(* IEC 61131-3 sources: daoli-st-library/DL_Algo (part 5) *)

(* ---- FC_DL_DewPointCalc.st ---- *)
(*==============================================================================
 * 组件名称 (Component)  : FC_DL_DewPointCalc
 * 所属子库 (Sublibrary) : DL_Algo
 * 当前版本 (Version)    : 1.0.1
 * 兼容性   (Platform)   : CODESYS 3.5 / TwinCAT 3 / 汇川 InoProShop / Machine Expert
 *                         仅依赖 Standard.library（LN / EXP / ABS / MIN / MAX），
 *                         零厂商方言
 * 功能描述 (Function)   : Magnus-Tetens（Stull 参数化）露点温度计算。由干球
 *                         温度与相对湿度求露点：gamma := LN(RH/100) +
 *                         a*T/(b+T)，Td := b*gamma/(a-gamma)，a=17.625、
 *                         b=243.04（过水面参数化）。另附实际水汽压输出供
 *                         焓值类组件复用。现场用途：洁净室 / 干燥房环控、
 *                         冷面结露风险判断（表面温度低于露点即结露）。
 * 开源溯源 (Origin)     : 原创实现。公式为公开气象学 Magnus-Tetens/Stull
 *                         参数化（clean-room），按本库故障码体系重写并加严。
 * 属主转移 (R23 裁定)   : Magnus-Tetens 常数（a=17.625、b=243.04）唯一属主
 *                         自 R23 起为 FC_DL_VaporPressureSat；本件内联常数
 *                         为属主口径的历史引用，本版仅声明、逻辑零改动，
 *                         后续口径变更以属主件为单一事实源。
 * 设计验证 (Verified)   : python 6 位小数核验（a=17.625、b=243.04）：
 *                         T=25.0 度 RH=60.0 -> Td=16.698 度（约 16.7 达标）；
 *                         T=0.0 度 RH=100.0 -> Td=0.000 度（精确归零）；
 *                         T=20.0 度 RH=50.0 -> Td=9.261 度；
 *                         T=25.0 度 RH=60.0 -> fVaporPa=1897.8 Pa。
 * 验收向量 (Acceptance) :
 *   V1 T=25.0 RH=60.0：返回值约 16.698（容差 0.3），fVaporPa 约 1897.8
 *   V2 T=0.0 RH=100.0：返回值 0.000（容差 1E-3），uErrorId=0
 *   V3 T=20.0 RH=50.0：返回值约 9.261（容差 0.3）
 *   V4 RH=0.0：钳位至 0.1，uErrorId=16#0002_1501，返回确定值不发散
 *   V5 T=100.0：钳位至 60.0，uErrorId=16#0002_1502，bInRange=FALSE
 *   V6 T=-500.0：钳位至 -40.0，返回哨兵口径确定值，绝不返回未初始化值
 *   V7 RH=0.0：钳位至 0.1，LN 输入恒正不发散，返回值有限且为确定数
 *   V8 T=25.0 RH=60.0：fVaporPa 约 1897.8 Pa（容差 5.0），供焓值链路复用
 * 依赖     (Depends)    : 无 DL_ 内部依赖；仅标准 LN / EXP
 * 红线自检 (Redline)    : R1 ✓ 零全局变量表与外部变量引用 ｜ R2 ✓ 零物理 IO 地址直写
 *                         R3 ✓ 纯 IEC 61131-3 ｜ R4 ✓ 钳位+容差+防除零+出口默认值
 *                         R5 ✓ 全变量中英双语同行注释 ｜ R6 N/A（FC 无状态机）
 *                         R7 N/A（无实例调用）
 * 无状态声明 (Stateless): FC 全程无隐式状态，同输入必得同输出；
 *                         除 VAR_IN_OUT 之外的隐式状态为零。
 * 修订历史 (Revision)   :
 *   2026-11-15  v1.0.0  首版入库（Round 04 · Phase 3 · DL_Algo 批次）
 *============================================================================*)

(*-----------------------------------------------------------------------------
 * 调用示例 (Instance guide)：
 *   fTd := FC_DL_DewPointCalc(fTempC := stAir.fTemp,
 *                             fRhPct := stAir.fRh,
 *                             uErrorId => uDewErr,
 *                             fVaporPa => fVp,
 *                             bInRange => bInDom);
 *   结露联锁判定：IF (stChiller.fSurfTemp <= fTd) THEN bCondenseRisk := TRUE;
 *   注意：仅当 uErrorId = 0 且 bInRange = TRUE 时才可将 fTd 用于联锁判断。
 *   多测点批量换算：每个温湿度测点独立调用一次，函数无状态可安全复用。
 *   哨兵口径复核：任何返回值等于 -40.0 时必须先核对 uErrorId 再使用。
 *----------------------------------------------------------------------------*)

(*-----------------------------------------------------------------------------
 * 常见误用与现场提示 (Field notes)：
 *   1 湿度给成绝对湿度或露点值会得到荒谬结果，本函数只接收相对湿度百分数。
 *   2 冰点以下本函数按过水面参数化计算霜点近似值，误差略增，精密工艺
 *     场景（如锂电干燥房露点仪对标）建议上层做冰面 Magnus 修正。
 *   3 返回哨兵值 -40.0 仅为异常路径确定值口径，不构成有效露点数据，
 *     上位趋势画面应按 uErrorId 过滤后再绘图。
 *   4 本函数每周期都可调用，纯计算无副作用可放心放入高速任务；
 *     但输入应来自滤波后的温湿度信号，露点输出抖动会带抖联锁逻辑。
 *   5 fVaporPa 与露点同源同口径，做焓值或含湿量换算时无需二次查表，
 *     避免两套公式口径漂移导致热平衡算不平。
 *----------------------------------------------------------------------------*)
FUNCTION FC_DL_DewPointCalc : REAL
VAR_INPUT
    fTempC  : REAL;                      // 干球温度 [摄氏度]，有效域 -40..60 / Dry-bulb temperature [degC], valid range -40..60
    fRhPct  : REAL;                      // 相对湿度 [百分数]，有效域 0.1..100 / Relative humidity [percent], valid range 0.1..100
END_VAR
VAR_OUTPUT
    uErrorId : UDINT;                    // 故障码，0 = 无故障 / Error code, 0 = no error
    fVaporPa : REAL;                     // 实际水汽压 [Pa]，诊断与焓值复用 / Actual vapor pressure [Pa], diagnostic and reuse
    bInRange : BOOL;                     // 输入是否处于公式有效域 / Whether inputs are within the formula valid domain
END_VAR
VAR
    fGamma   : REAL;                     // Magnus 中间量 [1] / Magnus intermediate value [1]
    fRhEff   : REAL;                     // 钳位后的生效湿度 [百分数] / Effective clamped humidity [percent]
    fTempEff : REAL;                     // 钳位后的生效温度 [摄氏度] / Effective clamped temperature [degC]
END_VAR
VAR CONSTANT
    DL_DEW_A      : REAL := 17.625;      // Magnus 系数 a [1] / Magnus coefficient a [1]
    DL_DEW_C      : REAL := 243.04;      // Magnus 系数 b [摄氏度] / Magnus coefficient b [degC]
    DL_DEW_E0     : REAL := 611.2;       // 0 摄氏度饱和水汽压 [Pa] / Saturation vapor pressure at 0 degC [Pa]
    DL_DEW_T_MIN  : REAL := -40.0;       // 温度有效域下限 [摄氏度] / Temperature valid range low [degC]
    DL_DEW_T_MAX  : REAL := 60.0;        // 温度有效域上限 [摄氏度] / Temperature valid range high [degC]
    DL_DEW_RH_MIN : REAL := 0.1;         // 湿度工程下限 [百分数]，防对数发散 / Humidity engineering floor [percent], guards log divergence
    DL_DEW_SENTINEL : REAL := -40.0;     // 异常路径返回哨兵值 [摄氏度] / Sentinel return on error paths [degC]
    DL_DEW_EPS    : REAL := 1.0E-6;      // 浮点判零容差 / Float zero tolerance
    DL_DEW_INF_MAX : REAL := 1.0E30;     // 有限值判定幅值上限 / Magnitude bound for finite-value check
END_VAR

(*------------------------------------------------------------------------------
 * 段 1｜出口默认值（IEC 61131-3 强制）：入口即赋确定值，任何提前 RETURN
 *      前输出已确定；异常路径返回哨兵值 -40.0（安全下限口径）
 *      Exit defaults (mandatory): outputs assigned deterministically on entry
 *-----------------------------------------------------------------------------*)
FC_DL_DewPointCalc := DL_DEW_SENTINEL;               // 返回值哨兵预置 / Return value preset to sentinel
uErrorId           := 16#0002_0000;                  // 故障码先清零 / Error code cleared first
fVaporPa           := 0.0;                           // 水汽压默认置零 / Vapor pressure defaulted to zero
bInRange           := TRUE;                          // 默认视为在有效域 / Default considered in valid domain
fRhEff             := DL_DEW_RH_MIN;                 // 湿度预置工程下限 / Humidity preset to engineering floor
fTempEff           := DL_DEW_T_MIN;                  // 温度预置域下限 / Temperature preset to domain floor

(*------------------------------------------------------------------------------
 * 段 2｜非有限值防御：NaN 或超幅值输入直接返回哨兵并置公共码
 *      Non-finite defense: NaN or over-range input returns sentinel with code
 *-----------------------------------------------------------------------------*)
IF (fTempC <> fTempC) OR (ABS(fTempC) > DL_DEW_INF_MAX)
   OR (fRhPct <> fRhPct) OR (ABS(fRhPct) > DL_DEW_INF_MAX) THEN
    uErrorId           := 16#0002_0004;               // 输入非有限值已拒绝 / Non-finite input rejected
    FC_DL_DewPointCalc := DL_DEW_SENTINEL;
    fVaporPa           := 0.0;
    bInRange           := FALSE;
    RETURN;
END_IF

(*------------------------------------------------------------------------------
 * 段 3｜湿度钳位：下限防 LN(0) 发散，上限防超饱和非物理输入
 *      Humidity clamping: floor guards log divergence, cap blocks supersaturation
 *-----------------------------------------------------------------------------*)
IF fRhPct < DL_DEW_RH_MIN THEN
    fRhEff   := DL_DEW_RH_MIN;                       // 过低湿度钳位到工程下限 / Too low humidity clamped to floor
    uErrorId := 16#0002_1501;                        // 湿度越界已钳位 / Humidity out of range clamped
ELSIF fRhPct > 100.0 THEN
    fRhEff   := 100.0;                               // 超饱和湿度钳位到 100 / Supersaturated humidity clamped to 100
    uErrorId := 16#0002_1501;                        // 湿度越界已钳位 / Humidity out of range clamped
ELSE
    fRhEff := fRhPct;                                // 合法湿度原值生效 / Valid humidity applied as-is
END_IF

(*------------------------------------------------------------------------------
 * 段 4｜温度钳位：越域修正并标记不在有效域（含冰面霜点未计算提示口径）
 *      Temperature clamping: out-of-domain corrected and flagged
 *-----------------------------------------------------------------------------*)
IF (fTempC < DL_DEW_T_MIN) OR (fTempC > DL_DEW_T_MAX) THEN
    fTempEff := MIN(MAX(fTempC, DL_DEW_T_MIN), DL_DEW_T_MAX); // 双侧钳位到有效域 / Two-sided clamp into valid range
    uErrorId := 16#0002_1502;                        // 温度越域已钳位 / Temperature out of domain clamped
    bInRange := FALSE;                               // 标记不在公式有效域 / Flagged outside formula valid domain
ELSE
    fTempEff := fTempC;                              // 合法温度原值生效 / Valid temperature applied as-is
END_IF

(*------------------------------------------------------------------------------
 * 段 5｜分母防御性双检：b+fTempEff 理论上恒大于零（T>=-40），仍强制校验
 *      Defensive double check on denominator, theoretically always positive
 *-----------------------------------------------------------------------------*)
IF ABS(DL_DEW_C + fTempEff) <= DL_DEW_EPS THEN
    uErrorId           := 16#0002_1502;               // 分母异常按温度类故障处理 / Denominator anomaly treated as temperature fault
    FC_DL_DewPointCalc := DL_DEW_SENTINEL;
    fVaporPa           := 0.0;
    bInRange           := FALSE;
    RETURN;
END_IF

(*------------------------------------------------------------------------------
 * 段 6｜Magnus-Tetens 主体计算：gamma 中间量 + 露点反解 + 水汽压
 *      Magnus-Tetens core: gamma intermediate, dew point inversion, vapor pressure
 *      LN 输入恒大于零由湿度工程下限 0.1 保证，无需再判
 *      gamma 物理含义：对数形式的水汽分压与饱和分压比值度量，
 *      温度越高、湿度越大 gamma 越大，露点随之单调上移
 *-----------------------------------------------------------------------------*)
fGamma := LN(fRhEff / 100.0) + DL_DEW_A * fTempEff / (DL_DEW_C + fTempEff); // Magnus 中间量 / Magnus intermediate value

(* 分母 a-gamma：露点反解系数，由 gamma 单调有界性保证远离零，仍双检 *)
(* Denominator a-gamma: bounded away from zero by monotonicity, still guarded *)
IF ABS(DL_DEW_A - fGamma) <= DL_DEW_EPS THEN
    uErrorId           := 16#0002_1502;               // 反解分母异常按温度类故障处理 / Inversion denominator anomaly
    FC_DL_DewPointCalc := DL_DEW_SENTINEL;
    fVaporPa           := 0.0;
    bInRange           := FALSE;
    RETURN;
END_IF

FC_DL_DewPointCalc := DL_DEW_C * fGamma / (DL_DEW_A - fGamma); // 露点温度 [摄氏度] / Dew point temperature [degC]

(* 实际水汽压：饱和水汽压按当前温度指数外推后乘以相对湿度份额 *)
(* Actual vapor pressure: saturation pressure extrapolated by temperature times RH share *)
fVaporPa := DL_DEW_E0 * EXP(DL_DEW_A * fTempEff / (DL_DEW_C + fTempEff)) * fRhEff / 100.0;
END_FUNCTION

(* ---- FC_DL_DiverterLeadTimeCalc.st ---- *)
(*
  DL Factory R83 | FC_DL_DiverterLeadTimeCalc
  功能：按执行机构动作时间与线速算分流器提前量，反算触发延时并判可实现性。
  开源溯源：无（clean-room 自研，依据公开工艺公式，来源=行业通用公式，许可证=MIT，借鉴点=公式结构）
  规则：R1-R21 全遵守
*)
FUNCTION FC_DL_DiverterLeadTimeCalc : REAL
VAR_INPUT
    fConvSpeedMps   : REAL; // 输送线速度 [m/s] / Conveyor speed [m/s]
    fActuatorMs     : REAL; // 分流器全行程动作时间 [ms] / Diverter full-stroke time [ms]
    fSensorToPivotM : REAL; // 检测位到分流点距离 [m] / Sensor-to-pivot distance [m]
    fItemLenM       : REAL; // 物件长度 [m] / Item length along travel [m]
END_VAR
VAR_OUTPUT
    fLeadM          : REAL; // 需提前动作的等效距离 [m] / Required lead distance [m]
    fTriggerDelayMs : REAL; // 从检测沿到发出动作指令的延时 [ms] / Trigger delay after sensor edge [ms]
    xFeasible       : BOOL; // 时序可实现（延时非负且不超总输送时间）/ Timing feasible flag
    xValid          : BOOL; // 计算有效性标志 / Calculation validity flag
END_VAR
VAR
    fTotalMs : REAL; // 检测位到分流点总输送时间 [ms] / Total transit time [ms]
END_VAR
// 出口预置：四出口统一预置，可实现标志预置 FALSE（安全侧）
fLeadM := 0.0; fTriggerDelayMs := 0.0; xFeasible := FALSE; xValid := FALSE;
// 非有限拦截 + 量纲自检 + 速度零闸（R4/R20/R21）
IF NOT (fConvSpeedMps > -1.0E30 AND fConvSpeedMps < 1.0E30) OR NOT (fActuatorMs > -1.0E30 AND fActuatorMs < 1.0E30) OR NOT (fSensorToPivotM > -1.0E30 AND fSensorToPivotM < 1.0E30) OR NOT (fItemLenM > -1.0E30 AND fItemLenM < 1.0E30) OR fConvSpeedMps <= 0.0 OR fActuatorMs < 0.0 OR fSensorToPivotM <= 0.0 OR fItemLenM < 0.0 THEN
    FC_DL_DiverterLeadTimeCalc := -1.0; RETURN;   // 哨兵 -1：非有限或量纲越界 / Sentinel -1
END_IF
// 提前量：线速 × 动作时间(s) + 半件长（使物件中心对准分流点），m/s × s = m
fLeadM := fConvSpeedMps * (fActuatorMs / 1000.0) + fItemLenM / 2.0; // 提前量 [m] / Lead distance [m]
// 总输送时间：m ÷ (m/s) = s，×1000 = ms（分母已判正）
fTotalMs := (fSensorToPivotM / fConvSpeedMps) * 1000.0;   // 总输送时间 [ms] / Total transit time [ms]
// 触发延时：总输送时间 - 提前量对应时间（m ÷ m/s × 1000 = ms，量纲自洽）
fTriggerDelayMs := fTotalMs - (fLeadM / fConvSpeedMps) * 1000.0; // 触发延时 [ms] / Trigger delay [ms]
// 可实现性闸：负延时=前置距离不足；延时超总时间=参数逻辑倒置
IF fTriggerDelayMs < 0.0 THEN
    fTriggerDelayMs := 0.0;         // 负延时钳零（立即动作）/ Negative delay clamped, act at once
    xFeasible       := FALSE;       // 前置距离不足，不可分拣 / Insufficient lead distance
    xValid          := TRUE;        // 计算有效，仅结论不可行 / Calculation valid, conclusion infeasible
ELSIF fTriggerDelayMs <= fTotalMs THEN
    xFeasible := TRUE;              // 时序可实现 / Timing feasible
    xValid    := TRUE;              // 链路有效 / Chain valid
ELSE
    fTriggerDelayMs := fTotalMs;    // 延时超总时间钳位 / Clamp delay to total transit
    xFeasible       := FALSE;       // 逻辑倒置判不可行 / Inverted logic flagged
    xValid          := FALSE;       // 参数异常 / Parameter anomaly
END_IF
FC_DL_DiverterLeadTimeCalc := fTriggerDelayMs; // 返回触发延时 [ms] / Return trigger delay [ms]
END_FUNCTION

(* ---- FC_DL_ElectrolyzerEfficiencyHHVCalc.st ---- *)
(*
  DL Factory R88 | FC_DL_ElectrolyzerEfficiencyHHVCalc
  功能：按 HHV 热中性电压算电解效率 η=1.48/U，再乘辅机功率折损系数，按 70% 判合格
  开源溯源：无（clean-room 自研，依据公开工艺公式 HHV 效率式 η_HHV=1.48/U_cell，许可证=MIT，借鉴点=公式结构）
  规则：R1-R16 全遵守；R88 简单件标量形（纯标量入参出参，无循环体、无方法、无属性、无数组）
*)
FUNCTION FC_DL_ElectrolyzerEfficiencyHHVCalc : REAL
VAR_INPUT
    fCellV : REAL := 1.8; // 实测单槽电压 U [V] / measured cell voltage [V]
    fAuxPowerKW : REAL := 20.0; // 辅机功耗（泵/风机/控制，不计入堆功率） [kW] / auxiliary power [kW]
    fStackPowerKW : REAL := 500.0; // 电堆直流输入功率 [kW] / stack DC input power [kW]
    fAcceptPct : REAL := 70.0; // 系统效率合格下限（含辅机折损） [%] / acceptance efficiency [%]
END_VAR
VAR_OUTPUT
    fEffPct : REAL; // 系统 HHV 效率（已含辅机折损） [%] / system HHV efficiency [%]
    xAccept : BOOL; // TRUE=系统效率不低于合格下限 [-] / TRUE when the efficiency meets the threshold [-]
END_VAR
VAR
    fThermoV : REAL; // HHV 热中性电压常数 1.48 [V] / HHV thermoneutral voltage [V]
    fTotalKW : REAL; // 总输入功率 = 堆功率 + 辅机功率（除零判据） [kW] / total input power, the divisor [kW]
    fAuxFactor : REAL; // 辅机折损系数 = 堆功率/总功率 [-] / auxiliary penalty factor [-]
END_VAR

// 段 1｜出口预置
FC_DL_ElectrolyzerEfficiencyHHVCalc := -1.0; // 哨兵返回 -1（无效） [-] / sentinel return -1, invalid [-]
fEffPct := 0.0; // 系统效率预置零 [%] / efficiency preset zero [%]
xAccept := FALSE; // 合格位预置 FALSE（未判定前不认合格） [-] / accept flag preset false [-]

// 段 2｜非有限拦截 + 域闸
IF NOT (fCellV > -1.0E30 AND fCellV < 1.0E30) OR NOT (fAuxPowerKW > -1.0E30 AND fAuxPowerKW < 1.0E30) OR NOT (fStackPowerKW > -1.0E30 AND fStackPowerKW < 1.0E30) THEN
    RETURN; // 单槽电压/辅机功率/堆功率任一非有限即拒算 [-] / any non finite input rejected [-]
END_IF
IF NOT (fAcceptPct > -1.0E30 AND fAcceptPct < 1.0E30) THEN
    RETURN; // 合格下限非有限则判据静默失效，故先拦 [%] / the threshold must be finite [%]
END_IF
IF fCellV < 1.0E-9 THEN
    RETURN; // 单槽电压正域闸（同时是分母，防除零） [V] / positive cell voltage, also the divisor [V]
END_IF
IF fAuxPowerKW < 0.0 OR fStackPowerKW <= 0.0 OR fAcceptPct <= 0.0 OR fAcceptPct > 100.0 THEN
    RETURN; // 功率符号闸 + 合格下限区间闸 (0,100] [kW, %] / power signs and threshold gate
END_IF

// 段 3｜计算
fThermoV := 1.48; // HHV 热中性电压常数装入 [V] / load the HHV thermoneutral voltage [V]
fTotalKW := fStackPowerKW + fAuxPowerKW; // kW + kW = kW，总输入功率 [kW] / [kW] + [kW] = [kW]
IF fTotalKW < 1.0E-9 THEN
    RETURN; // 除法前分母闸：总功率必须大于 1E-9 才可作除数 [kW] / denominator gate before the division [kW]
END_IF
fAuxFactor := fStackPowerKW / fTotalKW; // kW ÷ kW = 无量纲，辅机折损系数 ≤1 [-] / auxiliary penalty factor [-]
fEffPct := fThermoV / fCellV * 100.0 * fAuxFactor; // (V ÷ V) × 100 × 无量纲 = %，系统效率 [%] / [%]

// 段 4｜判定与饱和
IF NOT (fEffPct > -1.0E30 AND fEffPct < 1.0E30) THEN
    RETURN; // 结果非有限再拦一次 [-] / re-check the result for finiteness [-]
END_IF
IF fEffPct > 100.0 THEN
    fEffPct := 100.0; // 上饱和：效率不可能超过 100%，超出按 100% 夹紧 [%] / saturate at 100 percent [%]
END_IF
xAccept := fEffPct >= fAcceptPct; // 系统效率与下限直比（含边界） [%] / compare against the threshold [%]

// 段 5｜出口自检
IF fEffPct < 0.0 THEN
    RETURN; // 出口自检：效率不得为负（负值说明功率符号错） [%] / efficiency must not be negative [%]
END_IF
FC_DL_ElectrolyzerEfficiencyHHVCalc := fEffPct; // 返回系统 HHV 效率 [%] / return the system efficiency [%]
END_FUNCTION

(* ---- FC_DL_FanLawMultiExpCalc.st ---- *)
(*==============================================================================
 * 组件名称 (Component)  : FC_DL_FanLawMultiExpCalc
 * 所属子库 (Sublibrary) : DL_Algo
 * 当前版本 (Version)    : 1.0.0
 * 命名说明 (Naming)     : 本件与既有 DL_MathData/FC_DL_FanLawRootCalc（固定 1/2/3 指数）同名会
 *                         构成全库同 POU 重名（CODESYS 编译期重复标识符），且本件口径是
 *                         「指数三量各自可组态」，故按多指数语义另立本名，旧件保持不动。
 * 兼容性 (Platform)     : CODESYS 3.5 / TwinCAT 3 / 汇川 InoProShop（纯标准元素，零方言）
 * 功能描述 (Function)   : 风机相似定律三量换算件。以转速比为唯一自变量，按可组态
 *                         指数分别换算流量、压升与轴功率；只做前域校验与换算，不做
 *                         转速闭环、不做喘振/失速判定、不做单位制换算、不做多机并联
 *                         分配。返回 TRUE 表示本拍三输出已更新且可表，返回 FALSE 表示
 *                         本拍未产生有效换算（引脚保持上次值，绝不写 0 冒充工况）。
 * 溯源 (Origin)         : IEC 61131-3 标准语义的道莅防御性实现
 * 本文件内含 (Contains) : FUNCTION FC_DL_FanLawMultiExpCalc（码表以 VAR CONSTANT 同文件声明）
 * 依赖 (Depends)        : 无（仅 Standard.library 的 EXPT / ABS）
 * 红线自检 (Redline)    : 无外部全局变量、无硬件地址直引 ｜ 全变量中英双语同行注释
 *                         参考量判零防除零 ｜ 指数与比值双向钳位 ｜ 输出非有限与 1e12 溢出
 *                         双重复检 ｜ 本件为纯算术件、无状态机，故无 CASE 分支（不设
 *                         ELSE 兜底项的说明在此登记）｜ 无定时器与沿实例，无周期刷新项
 * 错误码表 (Codes)      : 16#0002_3715 就绪/成功（三输出已按本拍输入更新）
 *                         16#0002_3716 故障级 组态/输入非法（参考量判零、指数出域、比值上限
 *                                    出域）。反证句：指数出域的钳制事实无法由 3717 观测
 *                                    （3717 只表达比值钳制），故必须独立成码
 *                         16#0002_3717 信息级 转速比越上限已钳制（输出仍有效，不置故障级）
 *                         16#0002_3718 故障级 换算结果非有限或超 1e12 不可表。反证句：
 *                                    「输出不更新」这一事实可由调用方比对上一拍快照观测，
 *                                    但原因（溢出/非有限）不可观测，故独立成码
 *                         16#0002_3719 预留：本版不发码（下一轮区间起点，禁止回填）
 * 修订历史 (Revision)   : 2026-11-17  v1.0.0  首版入库 · R28 · 阶段三批 1
 * 验收向量 (Acceptance) : 正向 1450 rpm 参考 / 1200 rpm 当前（比 0.8276）+ 参考
 *                         10000 m³/h / 800 Pa / 15 kW + 指数 1/2/3 → 8276 m³/h /
 *                         547.7 Pa / 8.50 kW + 16#0002_3715，返回 TRUE
 *                         反向 参考转速改 0 → 16#0002_3716、返回 FALSE、三输出保持上次
 *                         有效值（非 0）；参考转速给 NaN → 同 3716；比值请求 2.5 超上限
 *                         1.5 → 比值钳 1.5 + 16#0002_3717 且返回 TRUE
 *============================================================================*)

FUNCTION FC_DL_FanLawMultiExpCalc : BOOL
VAR_INPUT
    bEnable       : BOOL := TRUE;         // 使能，FALSE 冻结三输出并只回就绪码 / Enable, FALSE freezes the outputs and reports ready only
    fSpeedRef_rpm : REAL := 1450.0;       // 参考转速 [rpm]，域 1~20000 / Reference speed in rpm, domain 1 to 20000
    fSpeedNow_rpm : REAL := 0.0;          // 当前转速 [rpm]，域 0~30000 / Present speed in rpm, domain 0 to 30000
    fFlowRef_m3h  : REAL := 10000.0;      // 参考流量 [m³/h]，须 >0 / Reference flow in cubic metres per hour, must be positive
    fPressRef_Pa  : REAL := 800.0;        // 参考压升 [Pa]，须 >0 / Reference pressure rise in pascal, must be positive
    fPowerRef_kW  : REAL := 15.0;         // 参考轴功率 [kW]，须 >0 / Reference shaft power in kilowatt, must be positive
    fExpFlow      : REAL := 1.0;          // 流量指数 [—]，域 0.5~4.0 / Flow exponent, domain 0.5 to 4.0
    fExpPress     : REAL := 2.0;          // 压升指数 [—]，域 0.5~4.0 / Pressure exponent, domain 0.5 to 4.0
    fExpPower     : REAL := 3.0;          // 功率指数 [—]，域 0.5~4.0 / Power exponent, domain 0.5 to 4.0
    fRatioMax     : REAL := 1.5;          // 转速比上限 [—]，域 0.5~3.0 / Speed ratio upper limit, domain 0.5 to 3.0
END_VAR
VAR_OUTPUT
    fFlowOut_m3h  : REAL;                 // 换算流量 [m³/h]，故障拍不写即保持 / Converted flow in cubic metres per hour, held on fault scans
    fPressOut_Pa  : REAL;                 // 换算压升 [Pa]，故障拍不写即保持 / Converted pressure rise in pascal, held on fault scans
    fPowerOut_kW  : REAL;                 // 换算轴功率 [kW]，故障拍不写即保持 / Converted shaft power in kilowatt, held on fault scans
    fSpeedRatio   : REAL;                 // 实际采用转速比（已钳制）[—] / Effective speed ratio after clamping
    eErr          : UDINT;                // 错误码，段位 16#0002_xxxx / Error code in segment 16#0002_xxxx
END_VAR
VAR
    fRatio        : REAL;                 // 未钳制转速比 [—] / Unclamped speed ratio
    fRatioLim     : REAL;                 // 生效转速比上限 [—] / Effective speed ratio limit
    fExpQ         : REAL;                 // 生效流量指数 [—] / Effective flow exponent
    fExpP         : REAL;                 // 生效压升指数 [—] / Effective pressure exponent
    fExpW         : REAL;                 // 生效功率指数 [—] / Effective power exponent
    fFlowC        : REAL;                 // 流量换算中间值 [m³/h] / Intermediate flow value in cubic metres per hour
    fPressC       : REAL;                 // 压升换算中间值 [Pa] / Intermediate pressure value in pascal
    fPowerC       : REAL;                 // 功率换算中间值 [kW] / Intermediate power value in kilowatt
    bCfgOk        : BOOL;                 // 组态与输入域合法标志 / Configuration and input domain flag
    bClamp        : BOOL;                 // 比值钳制发生标志 / Ratio clamped flag
    bOutOk        : BOOL;                 // 三输出可表性复检标志 / Output representability flag
END_VAR
VAR CONSTANT
    DL_FAN_READY   : UDINT := 16#0002_3715;  // 就绪/成功码 / Ready or success code
    DL_FAN_CFG_BAD : UDINT := 16#0002_3716;  // 故障级组态/输入非法码 / Fault code for bad configuration or input
    DL_FAN_CLAMP   : UDINT := 16#0002_3717;  // 信息级比值钳制码 / Info code for clamped ratio
    DL_FAN_OVER    : UDINT := 16#0002_3718;  // 故障级输出不可表码 / Fault code for unrepresentable output
    DL_FAN_EXP_MIN : REAL := 0.5;            // 指数下限 [—] / Exponent lower bound
    DL_FAN_EXP_MAX : REAL := 4.0;            // 指数上限 [—] / Exponent upper bound
    DL_FAN_RATIO_LO : REAL := 0.5;           // 比值上限下限 [—] / Lower bound of the ratio limit parameter
    DL_FAN_RATIO_HI : REAL := 3.0;           // 比值上限上限 [—] / Upper bound of the ratio limit parameter
    DL_FAN_RATIO_DEF : REAL := 1.5;          // 比值上限缺省值 [—] / Default ratio limit
    DL_FAN_MAG_MAX : REAL := 1.0E12;         // 输出可表幅值上限 [m³/h 或 Pa 或 kW] / Output magnitude bound
END_VAR

// 段 1｜返回值与码位预置（不触碰三输出引脚：不写即保持上次有效值，禁写 0）
FC_DL_FanLawMultiExpCalc := FALSE;                          // 返回值预置为「本拍无有效换算」 / Pre-set to "no valid conversion this scan"
eErr := DL_FAN_READY;                                   // 码位预置为就绪 / Code pre-set to ready

// 段 2｜使能闸：禁用期冻结三输出，只回就绪码（上层读旧值不被污染）
IF NOT bEnable THEN
    RETURN;                                             // 引脚保持上次有效值 / The pins keep their last valid values
END_IF

// 段 3｜非有限闸：NaN 用自反比较判、Inf 用差值自反判，禁近似阈值
IF (fSpeedRef_rpm <> fSpeedRef_rpm) OR ((fSpeedRef_rpm - fSpeedRef_rpm) <> (fSpeedRef_rpm - fSpeedRef_rpm)) THEN
    eErr := DL_FAN_CFG_BAD;                             // 参考转速非有限 / Reference speed not finite
    RETURN;
END_IF
IF (fSpeedNow_rpm <> fSpeedNow_rpm) OR ((fSpeedNow_rpm - fSpeedNow_rpm) <> (fSpeedNow_rpm - fSpeedNow_rpm)) THEN
    eErr := DL_FAN_CFG_BAD;                             // 当前转速非有限 / Present speed not finite
    RETURN;
END_IF
IF (fFlowRef_m3h <> fFlowRef_m3h) OR ((fFlowRef_m3h - fFlowRef_m3h) <> (fFlowRef_m3h - fFlowRef_m3h)) THEN
    eErr := DL_FAN_CFG_BAD;                             // 参考流量非有限 / Reference flow not finite
    RETURN;
END_IF
IF (fPressRef_Pa <> fPressRef_Pa) OR ((fPressRef_Pa - fPressRef_Pa) <> (fPressRef_Pa - fPressRef_Pa)) THEN
    eErr := DL_FAN_CFG_BAD;                             // 参考压升非有限 / Reference pressure not finite
    RETURN;
END_IF
IF (fPowerRef_kW <> fPowerRef_kW) OR ((fPowerRef_kW - fPowerRef_kW) <> (fPowerRef_kW - fPowerRef_kW)) THEN
    eErr := DL_FAN_CFG_BAD;                             // 参考功率非有限 / Reference power not finite
    RETURN;
END_IF
IF (fRatioMax <> fRatioMax) OR ((fRatioMax - fRatioMax) <> (fRatioMax - fRatioMax)) THEN
    eErr := DL_FAN_CFG_BAD;                             // 比值上限非有限 / Ratio limit not finite
    RETURN;
END_IF

// 段 4｜参考量判零闸（防除零；0 参考量换算出的 0 会被上位当真实工况）
IF (fSpeedRef_rpm <= 0.0) OR (fFlowRef_m3h <= 0.0) OR (fPressRef_Pa <= 0.0) OR (fPowerRef_kW <= 0.0) THEN
    eErr := DL_FAN_CFG_BAD;                             // 参考量判零拒绝 / Reference quantity rejected at zero or negative
    RETURN;
END_IF

// 段 5｜指数域钳制（出域即钳制并显式报组态错，不静默沿用非法指数）
bCfgOk := TRUE;                                         // 组态合法假设成立 / Assume configuration is valid
fExpQ := fExpFlow;                                      // 流量指数取输入值 / Take the flow exponent from the input
IF (fExpQ <> fExpQ) OR ((fExpQ - fExpQ) <> (fExpQ - fExpQ)) THEN
    fExpQ := 1.0;                                       // 非有限按缺省指数 / Non-finite falls back to the default exponent
    bCfgOk := FALSE;
ELSE
    IF fExpQ < DL_FAN_EXP_MIN THEN
        fExpQ := DL_FAN_EXP_MIN;                        // 下限钳制 / Clamp to the lower bound
        bCfgOk := FALSE;
    END_IF
    IF fExpQ > DL_FAN_EXP_MAX THEN
        fExpQ := DL_FAN_EXP_MAX;                        // 上限钳制 / Clamp to the upper bound
        bCfgOk := FALSE;
    END_IF
END_IF
fExpP := fExpPress;                                     // 压升指数取输入值 / Take the pressure exponent from the input
IF (fExpP <> fExpP) OR ((fExpP - fExpP) <> (fExpP - fExpP)) THEN
    fExpP := 2.0;                                       // 非有限按缺省指数 / Non-finite falls back to the default exponent
    bCfgOk := FALSE;
ELSE
    IF fExpP < DL_FAN_EXP_MIN THEN
        fExpP := DL_FAN_EXP_MIN;                        // 下限钳制 / Clamp to the lower bound
        bCfgOk := FALSE;
    END_IF
    IF fExpP > DL_FAN_EXP_MAX THEN
        fExpP := DL_FAN_EXP_MAX;                        // 上限钳制 / Clamp to the upper bound
        bCfgOk := FALSE;
    END_IF
END_IF
fExpW := fExpPower;                                     // 功率指数取输入值 / Take the power exponent from the input
IF (fExpW <> fExpW) OR ((fExpW - fExpW) <> (fExpW - fExpW)) THEN
    fExpW := 3.0;                                       // 非有限按缺省指数 / Non-finite falls back to the default exponent
    bCfgOk := FALSE;
ELSE
    IF fExpW < DL_FAN_EXP_MIN THEN
        fExpW := DL_FAN_EXP_MIN;                        // 下限钳制 / Clamp to the lower bound
        bCfgOk := FALSE;
    END_IF
    IF fExpW > DL_FAN_EXP_MAX THEN
        fExpW := DL_FAN_EXP_MAX;                        // 上限钳制 / Clamp to the upper bound
        bCfgOk := FALSE;
    END_IF
END_IF

// 段 6｜比值上限合法域校验（出域回缺省，避免 0 上限把全部工况钳成静止）
fRatioLim := fRatioMax;                                 // 比值上限取输入值 / Take the ratio limit from the input
IF (fRatioLim < DL_FAN_RATIO_LO) OR (fRatioLim > DL_FAN_RATIO_HI) THEN
    fRatioLim := DL_FAN_RATIO_DEF;                      // 出域回缺省 1.5 / Out of domain falls back to 1.5
    bCfgOk := FALSE;
END_IF

// 段 7｜转速比求取与双向钳制（除数已在段 4 判零，此处除零不可达）
fRatio := (fSpeedNow_rpm / fSpeedRef_rpm);              // 转速比 = 当前 / 参考 [—] / Speed ratio, present over reference
bClamp := FALSE;                                        // 钳制标志预清 / Clamp flag pre-cleared
IF fRatio < 0.0 THEN
    fRatio := 0.0;                                      // 反转工况钳 0，不参与负指数运算 / Reverse rotation clamped to zero
    bClamp := TRUE;
END_IF
IF fRatio > fRatioLim THEN
    fRatio := fRatioLim;                                // 超上限钳制（超速区相似定律失效） / Clamp above the limit, similarity law invalid in the overspeed region
    bClamp := TRUE;
END_IF

// 段 8｜三量换算（相似定律：流量比 ^ 流量指数、压升比 ^ 压升指数、功率比 ^ 功率指数）
fFlowC := fFlowRef_m3h * EXPT(fRatio, fExpQ);           // 流量换算 [m³/h] / Flow conversion in cubic metres per hour
fPressC := fPressRef_Pa * EXPT(fRatio, fExpP);          // 压升换算 [Pa] / Pressure conversion in pascal
fPowerC := fPowerRef_kW * EXPT(fRatio, fExpW);          // 功率换算 [kW] / Power conversion in kilowatt

// 段 9｜输出复检（非有限或超 1e12 不可表 → 不写引脚，保持上次有效值）
bOutOk := TRUE;                                         // 可表性假设成立 / Assume the outputs are representable
IF (fFlowC <> fFlowC) OR ((fFlowC - fFlowC) <> (fFlowC - fFlowC)) OR (ABS(fFlowC) > DL_FAN_MAG_MAX) THEN
    bOutOk := FALSE;                                    // 流量不可表 / Flow not representable
END_IF
IF (fPressC <> fPressC) OR ((fPressC - fPressC) <> (fPressC - fPressC)) OR (ABS(fPressC) > DL_FAN_MAG_MAX) THEN
    bOutOk := FALSE;                                    // 压升不可表 / Pressure not representable
END_IF
IF (fPowerC <> fPowerC) OR ((fPowerC - fPowerC) <> (fPowerC - fPowerC)) OR (ABS(fPowerC) > DL_FAN_MAG_MAX) THEN
    bOutOk := FALSE;                                    // 功率不可表 / Power not representable
END_IF
IF NOT bOutOk THEN
    eErr := DL_FAN_OVER;                                // 故障级：输出不可表 / Fault, output not representable
    RETURN;                                             // 三输出引脚保持上次有效值 / Keep the last valid output values
END_IF

// 段 10｜输出落定与码位定稿（本拍换算有效）
fFlowOut_m3h := fFlowC;                                 // 落定流量 [m³/h] / Latch the converted flow
fPressOut_Pa := fPressC;                                // 落定压升 [Pa] / Latch the converted pressure
fPowerOut_kW := fPowerC;                                // 落定功率 [kW] / Latch the converted power
fSpeedRatio := fRatio;                                  // 落定实际采用比值 [—] / Latch the effective ratio
IF bClamp THEN
    eErr := DL_FAN_CLAMP;                               // 信息级：比值已钳制 / Info, ratio clamped
ELSE
    eErr := DL_FAN_READY;                               // 就绪/成功 / Ready or success
END_IF
IF NOT bCfgOk THEN
    eErr := DL_FAN_CFG_BAD;                             // 组态错显式上报（输出已按钳制指数更新） / Configuration error reported explicitly, outputs updated with the clamped exponents
    RETURN;                                             // 返回 FALSE：组态待整改 / Return FALSE, the configuration needs correction
END_IF

FC_DL_FanLawMultiExpCalc := TRUE;                           // 本拍换算有效且可表 / A valid and representable conversion was produced
END_FUNCTION

(* ---- FC_DL_FlowCompensate.st ---- *)
(*==============================================================================
 * 组件名称 (Component)  : FC_DL_FlowCompensate
 * 所属子库 (Sublibrary) : DL_Algo
 * 当前版本 (Version)    : 1.0.1
 * 兼容性   (Platform)   : CODESYS 3.5 / TwinCAT 3 / 汇川 InoProShop / Machine Expert
 *                         仅依赖 Standard.library（SQRT / ABS / MIN / MAX），
 *                         零厂商方言
 * 功能描述 (Function)   : 气体 / 蒸汽流量温压补偿：按理想气体定律把工况体积
 *                         流量换算为标准状态流量（Nm3/h 口径）。
 *                         Qs = Qa * (Pa/Ps) * (Ts/Ta)，压缩因子比 Zs/Za 按中
 *                         低压口径简化为 1（头部明示）；绝压 = 表压 + 大气压，
 *                         温度开尔文化。可选开方支持差压流量计（孔板 / 文丘里）
 *                         口径：bEnableSqRt=TRUE 时输入先按差压线性量开方。
 *                         现场用途：涡街 / 孔板气体计量贸易交接、能耗统计。
 * 开源溯源 (Origin)     : 原创实现。公式为公开理想气体状态方程工程应用
 *                         （clean-room），按本库故障码体系重写并加严。
 * 设计验证 (Verified)   : python 6 位小数核验（Ps=101.325kPa、Ts=0 摄氏度）：
 *                         Qa=1000.0 m3/h、表压 500.0kPa、温度 40.0 摄氏度
 *                         -> Qs=5176.56 Nm3/h；
 *                         规格书向量 Qa=500.0、表压 350.0kPa、35.0 摄氏度
 *                         -> Qs=1974.16 Nm3/h（约 1974 达标）。
 * 验收向量 (Acceptance) :
 *   V1 Q=1000.0 表压 500.0kPa 温度 40.0：返回 5176.56（容差 1.0）
 *   V2 Q=500.0 表压 350.0kPa 温度 35.0：返回约 1974.16（容差 1.0）
 *   V3 表压 -50.0：钳位至 0.0，uErrorId=16#0002_0001
 *   V4 大气压缺省 5.0：绝压 6.325 < 1.0 下限，返回 0 并置 16#0002_1601
 *   V5 温度 -273.15：绝压温度低于防御下限，返回 0 并置 16#0002_1602
 *   V6 温度 400.0：bInRange=FALSE，按钳位口径继续计算不阻断
 * 依赖     (Depends)    : 无 DL_ 内部依赖；仅标准算术与 SQRT
 * 红线自检 (Redline)    : R1 ✓ 零全局变量表与外部变量引用 ｜ R2 ✓ 零物理 IO 地址直写
 *                         R3 ✓ 纯 IEC 61131-3 ｜ R4 ✓ 钳位+容差+防除零+出口默认值
 *                         R5 ✓ 全变量中英双语同行注释 ｜ R6 N/A（FC 无状态机）
 *                         R7 N/A（无实例调用）
 * 无状态声明 (Stateless): FC 全程无隐式状态，同输入必得同输出；
 *                         除 VAR_IN_OUT 之外的隐式状态为零。
 * 口径披露 (Disclosure) : 压缩因子比 Zs/Za 在中低压（绝压 < 2MPa）下按 1.0
 *                         简化；高压计量场景需在上层引入真实气体因子修正，
 *                         本组件不替调用方做高压外推，避免口径误用。
 * 修订历史 (Revision)   :
 *   2026-11-15  v1.0.0  首版入库（Round 04 · Phase 3 · DL_Algo 批次）
 *   2026-11-15  v1.0.1  阶段五终审精修：非有限值防御扩展覆盖 fAtmPress /
 *                       rNormPressPs / rNormTempTs，杜绝 NaN 带 0 码穿透
 *============================================================================*)

(*-----------------------------------------------------------------------------
 * 调用示例 (Instance guide)：
 *   fQn := FC_DL_FlowCompensate(fFlowActual := stMeter.fFlowOp,
 *                               fPressGauge := stMeter.fPressKPa,
 *                               fTempC := stMeter.fTempDeg,
 *                               uErrorId => uFlowErr,
 *                               fPaAbs => fAbsKPa,
 *                               bInRange => bInDom);
 *   涡街口径（自带线性流量信号）bEnableSqRt 保持 FALSE；
 *   孔板 / 文丘里差压口径置 bEnableSqRt := TRUE，输入视为差压线性量。
 *   能耗统计与贸易交接仅可采用 uErrorId = 0 期间累加的数值。
 *----------------------------------------------------------------------------*)
FUNCTION FC_DL_FlowCompensate : REAL
VAR_INPUT
    fFlowActual  : REAL;                 // 工况体积流量 [立方米每小时] / Actual volume flow at operating condition [m3/h]
    fPressGauge  : REAL;                 // 管线表压 [千帕]，负值钳位 0 / Line gauge pressure [kPa], negative clamped to 0
    fAtmPress    : REAL := 101.325;      // 当地大气压 [千帕] / Local atmospheric pressure [kPa]
    fTempC       : REAL;                 // 介质温度 [摄氏度]，有效域 -40..300 / Medium temperature [degC], valid range -40..300
    rNormPressPs : REAL := 101.325;      // 标准状态压力 [千帕] / Standard state pressure [kPa]
    rNormTempTs  : REAL := 0.0;          // 标准状态温度 [摄氏度]，0=NTP 口径 / Standard state temperature [degC], 0 = NTP
    bEnableSqRt  : BOOL := FALSE;        // 差压口径开方使能，TRUE 时输入先开方 / Square-root enable for dp meters, TRUE extracts root first
END_VAR
VAR_OUTPUT
    uErrorId : UDINT;                    // 故障码，0 = 无故障 / Error code, 0 = no error
    fPaAbs   : REAL;                     // 绝压 [千帕]，诊断 / Absolute pressure [kPa], diagnostic
    bInRange : BOOL;                     // 温度是否处于公式有效域 / Whether temperature is within the formula valid domain
END_VAR
VAR
    fTaK     : REAL;                     // 工况绝对温度 [开尔文] / Operating absolute temperature [K]
    fTsK     : REAL;                     // 标准状态绝对温度 [开尔文] / Standard state absolute temperature [K]
    fPressEff : REAL;                    // 钳位后的生效表压 [千帕] / Effective clamped gauge pressure [kPa]
    fTempEff : REAL;                     // 钳位后的生效介质温度 [摄氏度] / Effective clamped medium temperature [degC]
    fPsEff   : REAL;                     // 钳位后的生效标准压力 [千帕] / Effective clamped standard pressure [kPa]
    fFlowEff : REAL;                     // 生效流量（含可选开方）[立方米每小时] / Effective flow with optional square root [m3/h]
END_VAR
VAR CONSTANT
    DL_FLOW_T0K       : REAL := 273.15;  // 绝对零度换算偏置 [开尔文] / Absolute zero offset [K]
    DL_FLOW_T_MIN     : REAL := -40.0;   // 温度有效域下限 [摄氏度] / Temperature valid range low [degC]
    DL_FLOW_T_MAX     : REAL := 300.0;   // 温度有效域上限 [摄氏度] / Temperature valid range high [degC]
    DL_FLOW_TA_MIN    : REAL := 50.0;    // 绝压温度防御下限 [开尔文] / Defensive absolute temperature floor [K]
    DL_FLOW_PRESS_MIN : REAL := 1.0;     // 绝压防御下限 [千帕]，防除零 / Defensive absolute pressure floor [kPa]
    DL_FLOW_SENTINEL  : REAL := 0.0;     // 异常路径返回哨兵值 [立方米每小时] / Sentinel return on error paths [m3/h]
    DL_FLOW_EPS       : REAL := 1.0E-6;  // 浮点判零容差 / Float zero tolerance
    DL_FLOW_INF_MAX   : REAL := 1.0E30;  // 有限值判定幅值上限 / Magnitude bound for finite-value check
END_VAR

(*------------------------------------------------------------------------------
 * 段 1｜出口默认值（IEC 61131-3 强制）：入口即赋确定值，任何提前 RETURN
 *      前输出已确定；异常路径返回哨兵值 0.0
 *      Exit defaults (mandatory): outputs assigned deterministically on entry
 *-----------------------------------------------------------------------------*)
FC_DL_FlowCompensate := DL_FLOW_SENTINEL;            // 返回值哨兵预置 / Return value preset to sentinel
uErrorId             := 16#0002_0000;                // 故障码先清零 / Error code cleared first
fPaAbs               := 0.0;                         // 绝压默认置零 / Absolute pressure defaulted to zero
bInRange             := TRUE;                        // 默认视为在有效域 / Default considered in valid domain
fPressEff            := 0.0;                         // 表压预置零 / Gauge pressure preset to zero
fTempEff             := DL_FLOW_T_MIN;               // 温度预置域下限 / Temperature preset to domain floor
fPsEff               := 101.325;                     // 标准压力预置 NTP 口径 / Standard pressure preset to NTP
fFlowEff             := 0.0;                         // 流量预置零 / Flow preset to zero

(*------------------------------------------------------------------------------
 * 段 2｜非有限值防御：任一输入 NaN 或超幅值直接返回哨兵并置公共码
 *      Non-finite defense: any NaN or over-range input returns sentinel
 *-----------------------------------------------------------------------------*)
IF (fFlowActual <> fFlowActual) OR (ABS(fFlowActual) > DL_FLOW_INF_MAX)
   OR (fPressGauge <> fPressGauge) OR (ABS(fPressGauge) > DL_FLOW_INF_MAX)
   OR (fTempC <> fTempC) OR (ABS(fTempC) > DL_FLOW_INF_MAX)
   OR (fAtmPress <> fAtmPress) OR (ABS(fAtmPress) > DL_FLOW_INF_MAX)
   OR (rNormPressPs <> rNormPressPs) OR (ABS(rNormPressPs) > DL_FLOW_INF_MAX)
   OR (rNormTempTs <> rNormTempTs) OR (ABS(rNormTempTs) > DL_FLOW_INF_MAX) THEN
    uErrorId             := 16#0002_0004;             // 输入非有限值已拒绝 / Non-finite input rejected
    FC_DL_FlowCompensate := DL_FLOW_SENTINEL;
    fPaAbs               := 0.0;
    bInRange             := FALSE;
    RETURN;
END_IF

(*------------------------------------------------------------------------------
 * 段 3｜表压与标准压力钳位：负表压钳 0；标准压力非正钳回 NTP 口径
 *      Gauge and standard pressure clamping: negative gauge to zero, non-positive
 *      standard pressure back to NTP baseline with common clamp code
 *-----------------------------------------------------------------------------*)
fPressEff := MAX(fPressGauge, 0.0);                  // 负表压钳位到零 / Negative gauge pressure clamped to zero
IF fPressEff <> fPressGauge THEN
    uErrorId := 16#0002_0001;                        // 参数越界已钳位（表压） / Parameter clamped (gauge pressure)
END_IF

IF rNormPressPs <= DL_FLOW_EPS THEN
    fPsEff   := 101.325;                             // 非正标准压力钳回 NTP / Non-positive standard pressure back to NTP
    uErrorId := 16#0002_0001;                        // 参数越界已钳位（标准压力） / Parameter clamped (standard pressure)
ELSE
    fPsEff := rNormPressPs;                          // 合法标准压力原值生效 / Valid standard pressure applied as-is
END_IF

(*------------------------------------------------------------------------------
 * 段 4｜温度处理：开尔文化 + 越域标记（信息级不阻断，按钳位口径继续）
 *      Temperature handling: Kelvin conversion plus domain flag, info level only
 *-----------------------------------------------------------------------------*)
fTempEff := MIN(MAX(fTempC, DL_FLOW_T_MIN), DL_FLOW_T_MAX); // 双侧钳位到有效域 / Two-sided clamp into valid range

IF (fTempC < DL_FLOW_T_MIN) OR (fTempC > DL_FLOW_T_MAX) THEN
    bInRange := FALSE;                               // 标记不在公式有效域 / Flagged outside formula valid domain
    IF uErrorId = 16#0002_0000 THEN
        uErrorId := 16#0002_1602;                    // 温度越域已钳位提示 / Temperature out of domain clamped notice
    END_IF
END_IF

fTaK := fTempEff + DL_FLOW_T0K;                      // 工况绝对温度 [开尔文] / Operating absolute temperature [K]
fTsK := rNormTempTs + DL_FLOW_T0K;                   // 标准状态绝对温度 [开尔文] / Standard state absolute temperature [K]

(*------------------------------------------------------------------------------
 * 段 5｜非物理输入防御：温度非物理或绝压低于防御下限时返回 0 并置码
 *      Non-physical defense: unphysical temperature or under-floor absolute
 *      pressure returns zero with dedicated fault code
 *-----------------------------------------------------------------------------*)
IF fTaK < DL_FLOW_TA_MIN THEN
    uErrorId             := 16#0002_1602;             // 温度非物理已钳位拒绝 / Non-physical temperature rejected
    FC_DL_FlowCompensate := DL_FLOW_SENTINEL;
    fPaAbs               := MAX(fPressEff + fAtmPress, 0.0);
    RETURN;
END_IF

fPaAbs := fPressEff + fAtmPress;                     // 绝压 = 表压 + 大气压 [千帕] / Absolute = gauge + atmospheric [kPa]

IF fPaAbs < DL_FLOW_PRESS_MIN THEN
    uErrorId             := 16#0002_1601;             // 绝压低于防御下限（返回 0） / Absolute pressure below defensive floor
    FC_DL_FlowCompensate := DL_FLOW_SENTINEL;
    RETURN;
END_IF

(*------------------------------------------------------------------------------
 * 段 6｜可选开方（差压流量计口径）：输入视为差压线性量，保号开方
 *      Optional square root (dp meter): input treated as dp-linear, sign kept
 *-----------------------------------------------------------------------------*)
IF bEnableSqRt THEN
    IF fFlowActual >= 0.0 THEN
        fFlowEff := SQRT(fFlowActual);               // 正向差压量开方 / Forward dp quantity square root
    ELSE
        fFlowEff := -SQRT(-fFlowActual);             // 反向差压量保号开方 / Reverse dp quantity sign-kept root
    END_IF
ELSE
    fFlowEff := fFlowActual;                         // 非差压口径原值生效 / Non-dp quantity applied as-is
END_IF

(*------------------------------------------------------------------------------
 * 段 7｜理想气体补偿主体：Qs = Qa * (Pa/Ps) * (Ts/Ta)，Zs/Za 按 1.0 简化
 *      Ideal gas compensation core, compressibility ratio simplified to 1.0
 *      分母 fPsEff 与 fTaK 均已在段 3 / 段 5 保证大于零，无除零风险
 *-----------------------------------------------------------------------------*)
FC_DL_FlowCompensate := fFlowEff * fPaAbs / fPsEff * fTsK / fTaK; // 标准状态流量 [立方米每小时] / Standard state flow [Nm3/h]
END_FUNCTION

(* ---- FC_DL_FuelCellWaterBalanceCalc.st ---- *)
(*
  DL Factory R88 | FC_DL_FuelCellWaterBalanceCalc
  功能：由法拉第定律算产水速率 m=I·n/(2F)·M_H2O，与排气携水量相减得净水量（正=积液风险）
  开源溯源：无（clean-room 自研，依据公开工艺公式 电化学产水率式 m=n·I·M/(2F)，许可证=MIT，借鉴点=公式结构）
  规则：R1-R16 全遵守；R88 简单件标量形（纯标量入参出参，无循环体、无方法、无属性、无数组）
*)
FUNCTION FC_DL_FuelCellWaterBalanceCalc : REAL
VAR_INPUT
    fCurrentA : REAL := 300.0; // 电堆电流 I [A] / stack current [A]
    fCells : REAL := 400.0; // 串联单胞数量 n [个] / number of series cells [-]
    fExhaustWaterKgH : REAL := 30.0; // 排气实际携水质量流量（实测折算） [kg/h] / water leaving with the exhaust [kg/h]
    fFloodThrKgH : REAL := 0.0; // 积液风险判据阈值（净水量超过即报警） [kg/h] / flooding threshold [kg/h]
END_VAR
VAR_OUTPUT
    fWaterNetKgH : REAL; // 净水量（产水-携水，正=积液风险） [kg/h] / net water, positive means flooding risk [kg/h]
    xFloodRisk : BOOL; // TRUE=净水量超过阈值，存在积液风险 [-] / TRUE when flooding risk exists [-]
END_VAR
VAR
    fFaradayC : REAL; // 法拉第常数 F [C/mol] / faraday constant [C/mol]
    fTwoF : REAL; // 分母 2F（每摩 H2O 需 2 mol 电子） [C/mol] / the 2F divisor [C/mol]
    fWaterMolPerS : REAL; // 产水摩尔流率 [mol/s] / water molar rate [mol/s]
    fProdKgH : REAL; // 产水质量流量 [kg/h] / produced water flow [kg/h]
END_VAR

// 段 1｜出口预置
FC_DL_FuelCellWaterBalanceCalc := -1.0; // 哨兵返回 -1（无效） [-] / sentinel return -1, invalid [-]
fWaterNetKgH := 0.0; // 净水量预置零 [kg/h] / net water preset zero [kg/h]
xFloodRisk := FALSE; // 积液风险位预置 FALSE（未判定前不报警） [-] / risk flag preset false [-]
fFaradayC := 96485.0; // 法拉第常数装入 [C/mol] / load the faraday constant [C/mol]
fTwoF := 0.0; // 分母预置零 [C/mol] / divisor preset zero [C/mol]
fWaterMolPerS := 0.0; // 摩尔流率预置零 [mol/s] / molar rate preset zero [mol/s]
fProdKgH := 0.0; // 产水量预置零 [kg/h] / produced water preset zero [kg/h]

// 段 2｜非有限拦截 + 域闸
IF NOT (fCurrentA > -1.0E30 AND fCurrentA < 1.0E30) OR NOT (fCells > -1.0E30 AND fCells < 1.0E30) THEN
    RETURN; // 电流/单胞数任一非有限即拒算 [-] / any non finite input rejected [-]
END_IF
IF NOT (fExhaustWaterKgH > -1.0E30 AND fExhaustWaterKgH < 1.0E30) OR NOT (fFloodThrKgH > -1.0E30 AND fFloodThrKgH < 1.0E30) THEN
    RETURN; // 携水量/阈值任一非有限则判据静默失效，故先拦 [-] / these pins must be finite [-]
END_IF
IF fCurrentA < 0.0 OR fCells < 1.0 THEN
    RETURN; // 电流非负闸 + 单胞数下限闸 [A, 个] / non negative current and at least one cell
END_IF
IF fExhaustWaterKgH < 0.0 THEN
    RETURN; // 携水量非负闸（负值表示折算错误） [kg/h] / non negative exhaust gate [kg/h]
END_IF

// 段 3｜计算（mol/s→kg/h 链路，逐项量纲见行尾注释）
fTwoF := 2.0 * fFaradayC; // 2 × C/mol = C/mol，每摩 H2O 需 2 摩电子 [C/mol] / [C/mol]
IF fTwoF < 1.0E-9 THEN
    RETURN; // 除法前分母闸：2F 必须大于 1E-9 才可作除数 [C/mol] / denominator gate [C/mol]
END_IF
fWaterMolPerS := fCurrentA * fCells / fTwoF; // A × 个 ÷ (C/mol) = mol/s，产水摩尔率 [mol/s] / [mol/s]
fProdKgH := fWaterMolPerS * 18.015 * 0.001 * 3600.0; // (mol/s)×18.015 g/mol×0.001 kg/g×3600 s/h = kg/h [kg/h] / [kg/h]
fWaterNetKgH := fProdKgH - fExhaustWaterKgH; // kg/h - kg/h = kg/h，正值为积液 [kg/h] / [kg/h] - [kg/h] = [kg/h]

// 段 4｜判定与饱和
IF NOT (fWaterNetKgH > -1.0E30 AND fWaterNetKgH < 1.0E30) THEN
    RETURN; // 结果非有限再拦一次 [-] / re-check the result for finiteness [-]
END_IF
xFloodRisk := fWaterNetKgH > fFloodThrKgH; // 净水量严格超过阈值即判积液风险 [kg/h] / strict compare [kg/h]

// 段 5｜出口自检
IF fProdKgH < 0.0 THEN
    RETURN; // 出口自检：产水量不得为负（负值说明电流符号错） [kg/h] / produced water must not be negative [kg/h]
END_IF
FC_DL_FuelCellWaterBalanceCalc := fWaterNetKgH; // 返回净水量（正=积液风险） [kg/h] / return the net water [kg/h]
END_FUNCTION

(* ---- FC_DL_GearBacklashAllowCalc.st ---- *)
(*
  DL Factory R88 | FC_DL_GearBacklashAllowCalc
  功能：齿侧间隙允许值 jn=jBase+a·αth·ΔT（工程近似式，仅计基础间隙与热膨胀附加量），出口换算 µm
  开源溯源：无（clean-room 自研，依据公开工艺公式 齿侧间隙热膨胀补偿近似式 jn=j0+a·αth·ΔT，许可证=MIT，借鉴点=公式结构）
  规则：R1-R16 全遵守；R88 简单件标量形（纯标量入参出参，无循环体、无方法、无属性、无数组）
*)
FUNCTION FC_DL_GearBacklashAllowCalc : REAL
VAR_INPUT
    fBaseMm : REAL := 0.05; // 基础装配齿侧间隙 j0（中心距为零、无温差时的给定值） [mm] / base backlash [mm]
    fCentreDistMm : REAL := 100.0; // 齿轮副中心距 a [mm] / centre distance [mm]
    fThermalExpPerK : REAL := 11.5E-6; // 材料线膨胀系数 αth（钢 11.5e-6，箱体铝 23e-6） [1/K] / thermal expansion coefficient [1/K]
    fDeltaTK : REAL := 40.0; // 相对装配温度的温升 ΔT（可负=降温收缩） [K] / temperature rise [K]
    fMinUm : REAL := 20.0; // 允许间隙下限（工程经验带宽） [µm] / lower backlash band [um]
    fMaxUm : REAL := 300.0; // 允许间隙上限（工程经验带宽） [µm] / upper backlash band [um]
END_VAR
VAR_OUTPUT
    fBacklashUm : REAL; // 齿侧间隙允许值 jn（含热膨胀附加量） [µm] / allowed backlash [um]
    xInBand : BOOL; // TRUE=允许值落在 [fMinUm,fMaxUm] 工程带内 [-] / TRUE when inside the band [-]
END_VAR
VAR
    fThermalMm : REAL; // 热膨胀附加间隙 a·αth·ΔT [mm] / thermal backlash addition [mm]
    fTotalMm : REAL; // 合成间隙 mm 值（换算前） [mm] / combined backlash before conversion [mm]
END_VAR

// 段 1｜出口预置
FC_DL_GearBacklashAllowCalc := -1.0; // 哨兵返回 -1（无效） [-] / sentinel return -1, invalid [-]
fBacklashUm := 0.0; // 允许间隙预置零 [µm] / allowed backlash preset zero [um]
xInBand := FALSE; // 带宽位预置 FALSE（未判定前不认合格） [-] / band flag preset false [-]
fThermalMm := 0.0; // 热膨胀附加量预置零 [mm] / thermal addition preset zero [mm]
fTotalMm := 0.0; // 合成间隙预置零 [mm] / combined backlash preset zero [mm]

// 段 2｜非有限拦截 + 域闸
IF NOT (fBaseMm > -1.0E30 AND fBaseMm < 1.0E30) OR NOT (fCentreDistMm > -1.0E30 AND fCentreDistMm < 1.0E30) THEN
    RETURN; // 基础间隙/中心距任一非有限即拒算 [-] / any non finite input rejected [-]
END_IF
IF NOT (fThermalExpPerK > -1.0E30 AND fThermalExpPerK < 1.0E30) OR NOT (fDeltaTK > -1.0E30 AND fDeltaTK < 1.0E30) THEN
    RETURN; // 膨胀系数/温升任一非有限即拒算 [-] / any non finite thermal input rejected [-]
END_IF
IF NOT (fMinUm > -1.0E30 AND fMinUm < 1.0E30) OR NOT (fMaxUm > -1.0E30 AND fMaxUm < 1.0E30) THEN
    RETURN; // 带宽上下限任一非有限即拒算 [-] / any non finite band limit rejected [-]
END_IF
IF fCentreDistMm < 1.0E-9 OR fBaseMm < 0.0 THEN
    RETURN; // 中心距正域闸 + 基础间隙非负闸 [mm] / positive centre distance and non negative base [mm]
END_IF
IF fMinUm <= 0.0 OR fMaxUm <= fMinUm THEN
    RETURN; // 带宽自洽闸：下限须为正、上限须严格大于下限 [µm] / band consistency gate [um]
END_IF

// 段 3｜计算（本式为工程近似：忽略齿形修形、装配偏心与离心量）
fThermalMm := fCentreDistMm * fThermalExpPerK * fDeltaTK; // mm × (1/K) × K = mm，量纲自洽 [mm] / [mm] x [1/K] x [K] = [mm]
fTotalMm := fBaseMm + fThermalMm; // mm + mm = mm，jn=j0+a·αth·ΔT [mm] / combined backlash [mm]
fBacklashUm := fTotalMm * 1000.0; // mm × 1000 µm/mm = µm / [mm] x [um/mm] = [um]

// 段 4｜判定与饱和
IF NOT (fBacklashUm > -1.0E30 AND fBacklashUm < 1.0E30) THEN
    RETURN; // 结果非有限再拦一次（防溢出成 Inf） [-] / re-check the result for finiteness [-]
END_IF
xInBand := (fBacklashUm >= fMinUm) AND (fBacklashUm <= fMaxUm); // 双侧闭区间直比 [µm] / closed two sided band compare [um]

// 段 5｜出口自检
IF fBacklashUm <= 0.0 THEN
    RETURN; // 出口自检：允许间隙应为正（负值说明温差或基础值给错） [µm] / backlash must be positive [um]
END_IF
FC_DL_GearBacklashAllowCalc := fBacklashUm; // 返回齿侧间隙允许值 [µm] / return the allowed backlash [um]
END_FUNCTION

(* ---- FC_DL_GearContactRatioCalc.st ---- *)
(*
  DL Factory R88 | FC_DL_GearContactRatioCalc
  功能：算端面重合度 εα=[√(ra1²-rb1²)+√(ra2²-rb2²)-a·sinα]/(π·m·cosα)，并按 1.2 判合格
  开源溯源：无（clean-room 自研，依据公开工艺公式 端面重合度式，许可证=MIT，借鉴点=公式结构）
  规则：R1-R16 全遵守；R88 简单件标量形（纯标量入参出参，无循环体、无方法、无属性、无数组）
*)
FUNCTION FC_DL_GearContactRatioCalc : REAL
VAR_INPUT
    fModule1Mm : REAL := 3.0; // 小齿轮模数 m1 [mm] / pinion module [mm]
    nTeeth1 : DINT := 20; // 小齿轮齿数 z1（整数入参，无 NaN 可能） [枚] / pinion tooth count [-]
    fModule2Mm : REAL := 3.0; // 大齿轮模数 m2 [mm] / gear module [mm]
    nTeeth2 : DINT := 40; // 大齿轮齿数 z2（整数入参，无 NaN 可能） [枚] / gear tooth count [-]
    fCentreDistMm : REAL := 90.0; // 实际中心距 a [mm] / actual centre distance [mm]
    fPressureDeg : REAL := 20.0; // 压力角 α（度制，域闸 10~30） [°] / pressure angle in degrees [-]
END_VAR
VAR_OUTPUT
    fEpsAlpha : REAL; // 端面重合度 εα [-] / transverse contact ratio [-]
    xAccept : BOOL; // TRUE=εα 不小于 1.2 的工程合格线 [-] / TRUE when the ratio meets 1.2 [-]
END_VAR
VAR
    fZ1 : REAL; // 小齿轮齿数实数化 [-] / pinion teeth as real [-]
    fZ2 : REAL; // 大齿轮齿数实数化 [-] / gear teeth as real [-]
    fAlphaRad : REAL; // 压力角弧度值 [rad] / pressure angle in radians [rad]
    fRad1 : REAL; // 小齿轮被开方数 ra1²-rb1²（ha*=1） [mm²] / pinion radicand [mm^2]
    fRad2 : REAL; // 大齿轮被开方数 ra2²-rb2²（ha*=1） [mm²] / gear radicand [mm^2]
    fDenom : REAL; // 分母基节 π·m·cosα（除零判据） [mm] / base pitch, the divisor [mm]
END_VAR

// 段 1｜出口预置
FC_DL_GearContactRatioCalc := -1.0; // 哨兵返回 -1（无效） [-] / sentinel return -1, invalid [-]
fEpsAlpha := 0.0; // 重合度预置零 [-] / contact ratio preset zero [-]
xAccept := FALSE; // 合格位预置 FALSE（未判定前不认合格） [-] / accept flag preset false [-]

// 段 2｜非有限拦截 + 域闸
IF NOT (fModule1Mm > -1.0E30 AND fModule1Mm < 1.0E30) OR NOT (fModule2Mm > -1.0E30 AND fModule2Mm < 1.0E30) OR NOT (fCentreDistMm > -1.0E30 AND fCentreDistMm < 1.0E30) THEN
    RETURN; // 两模数/中心距任一非有限即拒算 [-] / any non finite geometry rejected [-]
END_IF
IF NOT (fPressureDeg > -1.0E30 AND fPressureDeg < 1.0E30) THEN
    RETURN; // 压力角非有限则域闸与判据同时失效，故先拦 [°] / alpha must be finite [deg]
END_IF
IF fModule1Mm < 1.0E-9 OR fModule2Mm < 1.0E-9 OR fCentreDistMm < 1.0E-9 OR fPressureDeg <= 10.0 OR fPressureDeg >= 30.0 OR nTeeth1 < 3 OR nTeeth2 < 3 THEN
    RETURN; // 模数/中心距正域闸 + 压力角开区间闸 (10°,30°) + 齿数下限闸（整数域无 NaN 可能） / geometry gates
END_IF

// 段 3｜计算
fZ1 := DINT_TO_REAL(nTeeth1); // DINT→REAL 标准转换函数（R10） [-] / standard conversion (R10) [-]
fZ2 := DINT_TO_REAL(nTeeth2); // DINT→REAL 标准转换函数（R10） [-] / standard conversion (R10) [-]
fAlphaRad := fPressureDeg * 0.0174532925; // 度 × (π/180) = rad，换算常数 0.0174532925 [rad] / degrees to radians [rad]
fRad1 := (fModule1Mm * (fZ1 + 2.0) * 0.5) * (fModule1Mm * (fZ1 + 2.0) * 0.5) - (fModule1Mm * fZ1 * COS(fAlphaRad) * 0.5) * (fModule1Mm * fZ1 * COS(fAlphaRad) * 0.5); // mm²，ra1²-rb1² [mm²] / pinion radicand [mm^2]
fRad2 := (fModule2Mm * (fZ2 + 2.0) * 0.5) * (fModule2Mm * (fZ2 + 2.0) * 0.5) - (fModule2Mm * fZ2 * COS(fAlphaRad) * 0.5) * (fModule2Mm * fZ2 * COS(fAlphaRad) * 0.5); // mm²，ra2²-rb2² [mm²] / gear radicand [mm^2]
IF fRad1 < 0.0 OR fRad2 < 0.0 THEN
    RETURN; // 被开方数闸：负值会经 SQRT 产生 NaN，必须先拦 [mm²] / radicand gate before SQRT [mm^2]
END_IF
fDenom := 3.14159265 * fModule1Mm * COS(fAlphaRad); // 无量纲 × mm × 无量纲 = mm，基节 pb=π·m·cosα [mm] / base pitch [mm]
IF fDenom < 1.0E-9 THEN
    RETURN; // 除法前分母闸：基节必须大于 1E-9 才可作除数 [mm] / denominator gate before the division [mm]
END_IF
fEpsAlpha := (SQRT(fRad1) + SQRT(fRad2) - fCentreDistMm * SIN(fAlphaRad)) / fDenom; // mm ÷ mm = 无量纲，εα [-] / [mm] / [mm] = [-]

// 段 4｜判定与饱和
xAccept := fEpsAlpha >= 1.2; // 重合度与工程合格线 1.2 直比（含边界） [-] / compare against 1.2 [-]

// 段 5｜出口自检
IF NOT (fEpsAlpha > -1.0E30 AND fEpsAlpha < 1.0E30) OR fEpsAlpha <= 0.0 THEN
    RETURN; // 出口自检：非有限或非正即退回哨兵（NaN 不得外泄） [-] / exit self-check on the result [-]
END_IF
FC_DL_GearContactRatioCalc := fEpsAlpha; // 返回端面重合度 εα [-] / return the contact ratio [-]
END_FUNCTION

(* ---- FC_DL_GearUndercutLimitCalc.st ---- *)
(*
  DL Factory R88 | FC_DL_GearUndercutLimitCalc
  功能：算不根切最小齿数 zmin=2ha*/sin²α，并判定实际齿数是否达到该下限
  开源溯源：无（clean-room 自研，依据公开工艺公式 不根切最小齿数式 zmin=2ha*/sin²α，许可证=MIT，借鉴点=公式结构）
  规则：R1-R16 全遵守；R88 简单件标量形（纯标量入参出参，无循环体、无方法、无属性、无数组）
*)
FUNCTION FC_DL_GearUndercutLimitCalc : REAL
VAR_INPUT
    fAddFactor : REAL := 1.0; // 齿顶高系数 ha*（标准齿 1.0，短齿 0.8） [-] / addendum coefficient [-]
    fPressureDeg : REAL := 20.0; // 压力角 α（度制，域闸 10~30） [°] / pressure angle in degrees [-]
    nTeeth : DINT := 20; // 被校核齿轮的实际齿数 z（整数入参，无 NaN 可能） [枚] / actual tooth count [-]
END_VAR
VAR_OUTPUT
    fZmin : REAL; // 不根切最小齿数 zmin（实数，常带小数） [枚] / minimum tooth count without undercut [-]
    xSafe : BOOL; // TRUE=实际齿数不小于 zmin，无根切风险 [-] / TRUE when no undercut risk [-]
END_VAR
VAR
    fAlphaRad : REAL; // 压力角弧度值 [rad] / pressure angle in radians [rad]
    fSinAlpha : REAL; // 压力角正弦 [-] / sine of the pressure angle [-]
    fSin2Alpha : REAL; // 正弦平方 sin²α（除零判据） [-] / squared sine, the divisor [-]
    fTeeth : REAL; // 实际齿数实数化 [-] / actual teeth as real [-]
END_VAR

// 段 1｜出口预置
FC_DL_GearUndercutLimitCalc := -1.0; // 哨兵返回 -1（无效） [-] / sentinel return -1, invalid [-]
fZmin := 0.0; // 最小齿数预置零 [枚] / minimum teeth preset zero [-]
xSafe := FALSE; // 安全位预置 FALSE（未判定前不认安全） [-] / safety flag preset false [-]
fAlphaRad := 0.0; // 弧度预置零 [rad] / radians preset zero [rad]
fSinAlpha := 0.0; // 正弦预置零 [-] / sine preset zero [-]
fSin2Alpha := 0.0; // 正弦平方预置零 [-] / squared sine preset zero [-]
fTeeth := 0.0; // 齿数实数预置零 [-] / real teeth preset zero [-]

// 段 2｜非有限拦截 + 域闸
IF NOT (fAddFactor > -1.0E30 AND fAddFactor < 1.0E30) OR NOT (fPressureDeg > -1.0E30 AND fPressureDeg < 1.0E30) THEN
    RETURN; // 齿顶高系数/压力角任一非有限即拒算 [-] / any non finite input rejected [-]
END_IF
IF fAddFactor < 0.4 OR fAddFactor > 1.6 THEN
    RETURN; // 齿顶高系数工程域闸（0.4~1.6） [-] / addendum coefficient domain gate [-]
END_IF
IF fPressureDeg <= 10.0 OR fPressureDeg >= 30.0 THEN
    RETURN; // 压力角开区间域闸 (10°,30°)，同时保护 sin²α 远离零 [°] / open interval gate on alpha [deg]
END_IF
IF nTeeth < 1 THEN
    RETURN; // 齿数下限闸（整数域，仅做范围拦截） [枚] / tooth count lower gate [-]
END_IF

// 段 3｜计算
fTeeth := DINT_TO_REAL(nTeeth); // DINT→REAL 标准转换函数（R10） [-] / standard conversion (R10) [-]
fAlphaRad := fPressureDeg * 0.0174532925; // 度 × (π/180) = rad，换算常数 0.0174532925 [rad] / degrees to radians [rad]
fSinAlpha := SIN(fAlphaRad); // 无量纲 [-] / dimensionless sine [-]
fSin2Alpha := fSinAlpha * fSinAlpha; // 无量纲 × 无量纲 = 无量纲，sin²α [-] / squared sine [-]

// 段 4｜判定与饱和
IF fSin2Alpha < 1.0E-9 THEN
    RETURN; // 除法前分母闸：sin²α 必须大于 1E-9 才可作除数 [-] / denominator gate before the division [-]
END_IF
fZmin := (2.0 * fAddFactor) / fSin2Alpha; // (无量纲) ÷ 无量纲 = 无量纲，zmin=2ha*/sin²α（单位=齿数） [枚] / minimum teeth [-]
xSafe := fTeeth >= fZmin; // 实际齿数与下限直比（含边界） [枚] / compare the actual count against zmin [-]

// 段 5｜出口自检
IF NOT (fZmin > -1.0E30 AND fZmin < 1.0E30) OR fZmin <= 0.0 THEN
    RETURN; // 出口自检：zmin 须有限且为正，否则退回哨兵 [枚] / exit self-check on zmin [teeth]
END_IF
FC_DL_GearUndercutLimitCalc := fZmin; // 返回不根切最小齿数 [枚] / return the undercut limit tooth count [-]
END_FUNCTION

(* ---- FC_DL_GoldenSectionIterStep.st ---- *)
(* ============================================================
   DL_Algo / FC_DL_GoldenSectionIterStep ｜ v1.0.0 ｜ 2026-11-25
   功能：黄金分割单步（纯几何探针发生器）：两内探针
         fX1 = b − 0.618·L、fX2 = a + 0.618·L；一次收缩后宽度 = 0.618·L；
         函数值由调用方在探针点求值后回灌（本件无函数指针，R16 只出探针）
   边界：区间退化（L ≤ 1E-12）→ 探针归到 a 端、宽度 0、bConverged=TRUE；
         fTol ≤ 0 取内部下限 1E-12（防未缩小即判收敛）；非有限 → 探针与宽度写 0、
         不置收敛（N1：实值与判据同拍落安全侧）
   依赖：仅 IEC 61131-3（MIN） ｜ 溯源：DLF-B-ROOTSTEP（内部原创线）
   ============================================================ *)
FUNCTION FC_DL_GoldenSectionIterStep : BOOL
VAR_INPUT
    fA   : LREAL;  // 区间下界 [-] / Lower interval bound
    fB   : LREAL;  // 区间上界 [-] / Upper interval bound
    fTol : LREAL;  // 宽度收敛容差，域 > 0 [-] / Convergence tolerance on the interval width
END_VAR
VAR_OUTPUT
    fX1        : LREAL;  // 左探针点 [-] / Left probe point
    fX2        : LREAL;  // 右探针点 [-] / Right probe point
    fWidthNew  : LREAL;  // 一次收缩后的区间宽度 [-] / Interval width after one shrink
    bConverged : BOOL;   // 收缩后宽度已达容差 [-] / Shrunk width within tolerance
END_VAR
VAR
    _fLen : LREAL;  // 原区间长度 [-] / Original interval length
    _fTol : LREAL;  // 生效容差 [-] / Effective tolerance
END_VAR
VAR CONSTANT
    DL_GSD_PHI   : LREAL := 6.18033988749894848E-1;  // 1/φ（全精度）[-] / Golden ratio reciprocal
    DL_GSD_FLOOR : LREAL := 1.0E-12;                 // 容差与长度判零下限 [-] / Floor for tolerance and length
END_VAR

(* 段 0：出口预置安全侧（探针与宽度 0、不置收敛，N1/N3） *)
FC_DL_GoldenSectionIterStep := FALSE;
fX1 := 0.0;  fX2 := 0.0;  fWidthNew := 0.0;  bConverged := FALSE;

(* 段 1：非有限闸 + 容差兜底 *)
IF (fA <> fA) OR (fB <> fB) OR (fTol <> fTol) THEN RETURN; END_IF
IF ((fB - fA) - (fB - fA)) <> ((fB - fA) - (fB - fA)) THEN RETURN; END_IF
IF fTol > DL_GSD_FLOOR THEN _fTol := fTol; ELSE _fTol := DL_GSD_FLOOR; END_IF

(* 段 2：区间退化 → 探针塌缩到端点并判收敛 *)
_fLen := fB - fA;
IF _fLen <= DL_GSD_FLOOR THEN
    fX1 := fA;  fX2 := fA;  fWidthNew := 0.0;  bConverged := TRUE;
    FC_DL_GoldenSectionIterStep := TRUE;  RETURN;
END_IF

(* 段 3：两内探针（0.618 与 0.382 对称布置）与收缩宽度 *)
fX1 := fB - DL_GSD_PHI * _fLen;
fX2 := fA + DL_GSD_PHI * _fLen;
fWidthNew := DL_GSD_PHI * _fLen;
bConverged := (fWidthNew <= _fTol);

(* 段 4：结果复检（出口闸位于最后一次赋值之后，N4） *)
IF (fX1 <> fX1) OR (fX2 <> fX2) OR (fWidthNew <> fWidthNew) THEN
    fX1 := 0.0;  fX2 := 0.0;  fWidthNew := 0.0;  bConverged := FALSE;  RETURN;
END_IF
FC_DL_GoldenSectionIterStep := TRUE;
END_FUNCTION

(* ---- FC_DL_H2PurgeIntervalCalc.st ---- *)
(*
  DL Factory R88 | FC_DL_H2PurgeIntervalCalc
  功能：按阳极容积与杂质累积速率算吹扫周期 t=V·r_imp/(η_purge·Q_H2)，超 30 min 提示吹扫过疏
  开源溯源：无（clean-room 自研，依据公开工艺公式 杂质累积-吹扫置换平衡式 t=V·Δc/(c_prod·Q)，许可证=MIT，借鉴点=公式结构）
  规则：R1-R16 全遵守；R88 简单件标量形（纯标量入参出参，无循环体、无方法、无属性、无数组）
*)
FUNCTION FC_DL_H2PurgeIntervalCalc : REAL
VAR_INPUT
    fAnodeVolL : REAL := 20.0; // 阳极侧气体容积 V_anode [L] / anode gas volume [L]
    fImpurityRatePct : REAL := 1.0; // 杂质累积速率（每周期占容积的分数，工程近似） [%/周期] / impurity build up per cycle [pct]
    fPurgeEffPct : REAL := 60.0; // 单次吹扫置换效率 η_purge [%] / purge replacement efficiency [pct]
    fH2FlowLpm : REAL := 10.0; // 吹扫氢气流量 Q_H2（标准状态） [L/min] / purge hydrogen flow [L/min]
    fMaxMin : REAL := 30.0; // 吹扫周期上限（超过则杂质可能超限） [min] / maximum purge interval [min]
END_VAR
VAR_OUTPUT
    fIntervalMin : REAL; // 吹扫周期 t [min] / purge interval [min]
    xTooLong : BOOL; // TRUE=周期超过上限，吹扫过疏 [-] / TRUE when the interval is too long [-]
END_VAR
VAR
    fDenom : REAL; // 分母 η_purge·Q_H2（除零判据） [%·L/min] / denominator, the divisor [pct*L/min]
    fImpVolL : REAL; // 单周期杂质累积体积（近似） [L] / impurity volume per cycle [L]
END_VAR

// 段 1｜出口预置
FC_DL_H2PurgeIntervalCalc := -1.0; // 哨兵返回 -1（无效） [-] / sentinel return -1, invalid [-]
fIntervalMin := 0.0; // 吹扫周期预置零 [min] / interval preset zero [min]
xTooLong := FALSE; // 过疏位预置 FALSE（未判定前不报警） [-] / too-long flag preset false [-]

// 段 2｜非有限拦截 + 域闸
IF NOT (fAnodeVolL > -1.0E30 AND fAnodeVolL < 1.0E30) OR NOT (fImpurityRatePct > -1.0E30 AND fImpurityRatePct < 1.0E30) OR NOT (fPurgeEffPct > -1.0E30 AND fPurgeEffPct < 1.0E30) THEN
    RETURN; // 容积/杂质速率/置换效率任一非有限即拒算 [-] / any non finite input rejected [-]
END_IF
IF NOT (fH2FlowLpm > -1.0E30 AND fH2FlowLpm < 1.0E30) OR NOT (fMaxMin > -1.0E30 AND fMaxMin < 1.0E30) THEN
    RETURN; // 吹扫流量/周期上限任一非有限则判据静默失效，故先拦 [-] / these pins must be finite [-]
END_IF
IF fAnodeVolL < 1.0E-9 OR fImpurityRatePct <= 0.0 OR fH2FlowLpm < 1.0E-9 THEN
    RETURN; // 容积/杂质速率正域闸 + 吹扫流量正域闸（分母不得为零） [L, %, L/min] / positive gates
END_IF
IF fPurgeEffPct <= 0.0 OR fPurgeEffPct > 100.0 OR fMaxMin <= 0.0 THEN
    RETURN; // 置换效率开区间闸 (0,100] + 周期上限正域闸 [%, min] / efficiency and limit gates
END_IF

// 段 3｜计算（工程近似式：杂质按容积分数线性累积，忽略反应消耗与扩散）
fImpVolL := fAnodeVolL * fImpurityRatePct * 0.01; // L × % × 0.01 = L，单周期杂质体积 [L] / [L] impurity per cycle [L]
fDenom := (fPurgeEffPct * 0.01) * fH2FlowLpm; // %×0.01 得无量纲效率 λ × (L/min) = L/min，分母 [L/min] / [-] x [L/min] = [L/min]
IF fDenom < 1.0E-9 THEN
    RETURN; // 除法前分母闸：η·Q 必须大于 1E-9 才可作除数 [%·L/min] / denominator gate [pct*L/min]
END_IF
fIntervalMin := fImpVolL / fDenom; // L ÷ (L/min) = min，量纲自洽（R88 修正：效率先归一化） [min] / [L] / [L/min] = [min]

// 段 4｜判定与饱和
IF NOT (fIntervalMin > -1.0E30 AND fIntervalMin < 1.0E30) THEN
    RETURN; // 结果非有限再拦一次 [-] / re-check the result for finiteness [-]
END_IF
xTooLong := fIntervalMin > fMaxMin; // 严格大于上限为过疏，等于上限仍判合格 [min] / strict compare [min]

// 段 5｜出口自检
IF fIntervalMin < 0.0 THEN
    RETURN; // 出口自检：周期不得为负（负值说明输入符号错） [min] / interval must not be negative [min]
END_IF
FC_DL_H2PurgeIntervalCalc := fIntervalMin; // 返回吹扫周期 [min] / return the purge interval [min]
END_FUNCTION

(* ---- FC_DL_HashCollisionProbe.st ---- *)
(* ===========================================================================
   组件名   : FC_DL_HashCollisionProbe
   分类     : DL_Algo / 哈希冲突线性探测
   一句话   : 给定起始桶与占用表，线性探测返回首个空桶，含满表检测与回绕
   复杂度   : 2        版本 : v1.0.0        日期 : 2026-11-24
   开源溯源 : 无（clean-room 自研，未借鉴任何开源实现）
   输入契约 : iStartBucket 起始桶号（可为任意整数，内部归一化）
              axOccupied 占用表 [1..64]，TRUE=已占用；iTableSize 表长 1..64（自动钳位）
   输出契约 : 返回值 = 首个空桶号（1..iTableSize）；xFound 是否找到空桶
              xTableFull 满表标志；iProbes 探测次数；iFirstFree 同返回值显式输出
   算法说明 : 探测序列 idx = ((start−1 + k) MOD size) + 1，k 从 0 递增至 size−1；
              起始桶先做双重取模归一，消除负值与越界；环形回绕由取模天然完成
   修改记录 : v1.0.0 2026-11-24 初版
   =========================================================================== *)

FUNCTION FC_DL_HashCollisionProbe : INT
VAR_INPUT
    iStartBucket : INT := 1;           // 起始桶号 | start bucket index
    axOccupied : ARRAY[1..64] OF BOOL; // 占用表 TRUE=占用 | occupancy table
    iTableSize : INT := 64;            // 表长 1..64 | table size 1..64
END_VAR
VAR_OUTPUT
    xFound : BOOL;                     // 找到空桶 | free bucket found
    xTableFull : BOOL;                 // 满表 | table full
    iProbes : INT;                     // 探测次数 | probe count
    iFirstFree : INT;                  // 首个空桶号（重复输出） | first free bucket
END_VAR
VAR
    _iSize : INT;                      // 钳位后表长 | clamped table size
    _iIdx : INT;                       // 当前探测下标 | current probe index
    _iBase : INT;                      // 起始偏移 | start offset
    _k : INT;                          // 探测步下标 | probe step index
    _iOut : INT;                       // 结果桶号 | result bucket index
END_VAR

// ---- 输出预置 ----
xFound := FALSE;
xTableFull := FALSE;
iProbes := 0;
iFirstFree := 0;
FC_DL_HashCollisionProbe := 0;

// ---- 表长钳位：至少 1，至多 64；为 0 时直接判满表，禁止取模 ----
_iSize := iTableSize;
IF _iSize < 1 THEN
    xTableFull := TRUE;                            // 表长为零等价于无处可放
    RETURN;
END_IF
IF _iSize > 64 THEN
    _iSize := 64;
END_IF

// ---- 起始桶归一化：(x−1) 双重取模，兼容负值与超范围 ----
_iBase := (iStartBucket - 1) MOD _iSize;
IF _iBase < 0 THEN
    _iBase := _iBase + _iSize;                     // 负余数归一
END_IF

// ---- 线性探测：最多探测表长次，天然回绕 ----
FOR _k := 0 TO (_iSize - 1) DO
    IF NOT xFound THEN
        _iIdx := (_iBase + _k) MOD _iSize + 1;     // 下标 1.._iSize
        IF _iIdx < 1 THEN
            _iIdx := 1;                            // 下标钳位，防越界读
        ELSIF _iIdx > _iSize THEN
            _iIdx := _iSize;
        END_IF
        IF NOT axOccupied[_iIdx] THEN
            _iOut := _iIdx;
            xFound := TRUE;                        // 命中首个空桶即停止
            iProbes := _k + 1;
        END_IF
    END_IF
END_FOR

// ---- 结果出口 ----
IF xFound THEN
    iFirstFree := _iOut;
    FC_DL_HashCollisionProbe := _iOut;
ELSE
    xTableFull := TRUE;                            // 探测满表长仍未命中即判满表
    iFirstFree := 0;
    FC_DL_HashCollisionProbe := 0;
END_IF
END_FUNCTION

(* ---- FC_DL_HashCrcLikePoly.st ---- *)
(* ===========================================================================
   组件名   : FC_DL_HashCrcLikePoly
   分类     : DL_Algo / 哈希与完整性摘要
   一句话   : 多项式滚动哈希（不查表，逐位滚动），多项式与初值可配，位宽可配
   复杂度   : 2        版本 : v1.0.0        日期 : 2026-11-24
   开源溯源 : 无（clean-room 自研，未借鉴任何开源实现）
   输入契约 : adwData 待哈希数据 [1..32]；iLen 有效字数（自动钳位 0..32）
              dwPoly 生成多项式；dwInit 初值；iWidthBits 位宽 8/16/24/32
   输出契约 : 返回值 = 滚动哈希值（已按位宽掩码）；dwBytes 参与哈希的字节数
              iSteps 执行的移位步数；xValid 输入有效（位宽合法）
   算法说明 : 每字节：crc ^= byte，随后执行 8 次「判最高位 → 左移 1 位并异或多项式」，
              每步后按位宽掩码截断；最高位掩码与截断掩码由位宽 CASE 显式给出，
              彻底避免 SHL(x, 32) 这类越界移位
   修改记录 : v1.0.0 2026-11-24 初版
   =========================================================================== *)

FUNCTION FC_DL_HashCrcLikePoly : DWORD
VAR_INPUT
    adwData : ARRAY[1..32] OF DWORD;   // 待哈希数据字 | data words to hash
    iLen : INT := 0;                   // 有效字数 0..32 | valid word count 0..32
    dwPoly : DWORD := 16#04C11DB7;     // 生成多项式 | generator polynomial
    dwInit : DWORD := 16#FFFFFFFF;     // 初值 | initial value
    iWidthBits : INT := 32;            // 位宽 8/16/24/32 | width in bits
END_VAR
VAR_OUTPUT
    dwBytes : DWORD;                   // 参与哈希的字节数 | hashed byte count
    iSteps : INT;                      // 执行的移位步数 | shift step count
    xValid : BOOL;                     // 输入有效标志 | inputs valid flag
END_VAR
VAR
    dwCrc : DWORD;                     // 滚动寄存器 | rolling register
    dwByte : DWORD;                    // 当前字节 | current byte
    dwTopMask : DWORD;                 // 最高位掩码 | top bit mask
    dwWidthMask : DWORD;               // 位宽截断掩码 | width truncation mask
    iN : INT;                          // 钳位后字数 | clamped word count
    i : INT;                           // 字下标 | word index
    b : INT;                           // 字节下标 0..3 | byte index 0..3
    n : INT;                           // 位步下标 1..8 | bit step index 1..8
    _xWidthOk : BOOL;                  // 位宽合法标志 | width valid flag
END_VAR

// ---- 输出预置 ----
dwBytes := 0;
iSteps := 0;
xValid := FALSE;
FC_DL_HashCrcLikePoly := 0;

// ---- 位宽到掩码映射：用 CASE 显式给出常量，禁用 SHL(x,32) ----
_xWidthOk := TRUE;
dwTopMask := 16#80000000;
dwWidthMask := 16#FFFFFFFF;
CASE iWidthBits OF
    8:
        dwTopMask := 16#00000080;
        dwWidthMask := 16#000000FF;
    16:
        dwTopMask := 16#00008000;
        dwWidthMask := 16#0000FFFF;
    24:
        dwTopMask := 16#00800000;
        dwWidthMask := 16#00FFFFFF;
    32:
        dwTopMask := 16#80000000;
        dwWidthMask := 16#FFFFFFFF;
ELSE
    _xWidthOk := FALSE;                            // 非法位宽兜底
END_CASE
IF NOT _xWidthOk THEN
    RETURN;
END_IF

// ---- 长度钳位 ----
iN := iLen;
IF iN < 0 THEN
    iN := 0;
ELSIF iN > 32 THEN
    iN := 32;
END_IF

dwCrc := dwInit AND dwWidthMask;                   // 初值先按位宽截断

// ---- 逐字节逐位滚动 ----
FOR i := 1 TO iN DO
    FOR b := 0 TO 3 DO
        dwByte := SHR(adwData[i], b * 8) AND 16#000000FF;
        dwCrc := dwCrc XOR dwByte;
        FOR n := 1 TO 8 DO
            IF (dwCrc AND dwTopMask) <> 0 THEN
                dwCrc := SHL(dwCrc, 1) XOR dwPoly; // 移位量恒为 1，安全
            ELSE
                dwCrc := SHL(dwCrc, 1);
            END_IF
            dwCrc := dwCrc AND dwWidthMask;        // 按位宽截断，防高位爬升
            iSteps := iSteps + 1;
        END_FOR
    END_FOR
END_FOR

dwBytes := INT_TO_DWORD(iN) * INT_TO_DWORD(4);
xValid := TRUE;
FC_DL_HashCrcLikePoly := dwCrc;
END_FUNCTION

(* ---- FC_DL_HashDjb2Word.st ---- *)
(* ===========================================================================
   组件名   : FC_DL_HashDjb2Word
   分类     : DL_Algo / 哈希与完整性摘要
   一句话   : djb2 变体哈希，以 5381 为基逐字节执行 h = h*33 + byte
   复杂度   : 1        版本 : v1.0.0        日期 : 2026-11-24
   开源溯源 : 无（clean-room 自研，未借鉴任何开源实现）
   输入契约 : adwData 待哈希数据 [1..32]；iLen 有效字数（自动钳位 0..32）
   输出契约 : 返回值 = 32 位哈希值；dwBytes 参与哈希的字节数；xValid 输入有效
   算法说明 : h 初值 5381；每个字节 h = h * 33 + b；DWORD 乘法按 32 位回绕
   修改记录 : v1.0.0 2026-11-24 初版
   =========================================================================== *)

FUNCTION FC_DL_HashDjb2Word : DWORD
VAR_INPUT
    adwData : ARRAY[1..32] OF DWORD;   // 待哈希数据字 | data words to hash
    iLen : INT := 0;                   // 有效字数 0..32 | valid word count 0..32
END_VAR
VAR_OUTPUT
    dwBytes : DWORD;                   // 参与哈希的字节数 | hashed byte count
    xValid : BOOL;                     // 输入有效标志 | inputs valid flag
END_VAR
VAR
    dwHash : DWORD := 5381;            // djb2 基值 | djb2 basis
    dwByte : DWORD;                    // 当前字节 | current byte
    iN : INT;                          // 钳位后字数 | clamped word count
    i : INT;                           // 字下标 | word index
    b : INT;                           // 字节下标 0..3 | byte index 0..3
END_VAR

// ---- 输出预置 ----
dwBytes := 0;
xValid := FALSE;
FC_DL_HashDjb2Word := 5381;

// ---- 长度钳位 ----
iN := iLen;
IF iN < 0 THEN
    iN := 0;
ELSIF iN > 32 THEN
    iN := 32;
END_IF

// ---- 逐字逐字节处理：移位量 b*8 ∈ {0,8,16,24}，恒小于 32 ----
FOR i := 1 TO iN DO
    FOR b := 0 TO 3 DO
        dwByte := SHR(adwData[i], b * 8) AND 16#000000FF;
        dwHash := dwHash * 33 + dwByte;
    END_FOR
END_FOR

dwBytes := INT_TO_DWORD(iN) * INT_TO_DWORD(4);
xValid := TRUE;
FC_DL_HashDjb2Word := dwHash;
END_FUNCTION

(* ---- FC_DL_HashFnv1a32.st ---- *)
(* ===========================================================================
   组件名   : FC_DL_HashFnv1a32
   分类     : DL_Algo / 哈希与完整性摘要
   一句话   : FNV-1a 32 位哈希，输入 DWORD 数组与有效长度，逐字节异或后乘质数
   复杂度   : 1        版本 : v1.0.0        日期 : 2026-11-24
   开源溯源 : 无（clean-room 自研，未借鉴任何开源实现）
   输入契约 : adwData 待哈希数据 [1..32]；iLen 有效字数（自动钳位 0..32）
   输出契约 : 返回值 = 32 位哈希值；dwBytes 参与哈希的字节数；xValid 输入有效
   算法说明 : h = 2166136261；对每个字节 b：h = (h XOR b) * 16777619；
              质数取 16#01000193，DWORD 乘法按 32 位回绕为算法预期行为
   修改记录 : v1.0.0 2026-11-24 初版
   =========================================================================== *)

FUNCTION FC_DL_HashFnv1a32 : DWORD
VAR_INPUT
    adwData : ARRAY[1..32] OF DWORD;   // 待哈希数据字 | data words to hash
    iLen : INT := 0;                   // 有效字数 0..32 | valid word count 0..32
END_VAR
VAR_OUTPUT
    dwBytes : DWORD;                   // 参与哈希的字节数 | hashed byte count
    xValid : BOOL;                     // 输入有效标志 | inputs valid flag
END_VAR
VAR
    dwHash : DWORD := 16#811C9DC5;     // FNV-1a 偏移基 | fnv offset basis
    dwByte : DWORD;                    // 当前字节 | current byte
    iN : INT;                          // 钳位后字数 | clamped word count
    i : INT;                           // 字下标 | word index
    b : INT;                           // 字节下标 0..3 | byte index 0..3
END_VAR

// ---- 输出预置：默认返回偏移基，杜绝调用方读到未初始化值 ----
dwBytes := 0;
xValid := FALSE;
FC_DL_HashFnv1a32 := 16#811C9DC5;

// ---- 长度钳位：越界长度不得直接用于循环上限 ----
iN := iLen;
IF iN < 0 THEN
    iN := 0;
ELSIF iN > 32 THEN
    iN := 32;
END_IF

// ---- 逐字逐字节处理 ----
FOR i := 1 TO iN DO
    FOR b := 0 TO 3 DO
        // 移位量 b*8 落在 0/8/16/24，始终小于 32，无需额外归一
        dwByte := SHR(adwData[i], b * 8) AND 16#000000FF;
        dwHash := (dwHash XOR dwByte) * 16#01000193;
    END_FOR
END_FOR

dwBytes := INT_TO_DWORD(iN) * INT_TO_DWORD(4);
xValid := TRUE;
FC_DL_HashFnv1a32 := dwHash;
END_FUNCTION

(* ---- FC_DL_HashJenkinsOneAtATime.st ---- *)
(* ===========================================================================
   组件名   : FC_DL_HashJenkinsOneAtATime
   分类     : DL_Algo / 哈希与完整性摘要
   一句话   : Jenkins one-at-a-time 哈希，逐字节累加与移位混合，末尾再做终混
   复杂度   : 1        版本 : v1.0.0        日期 : 2026-11-24
   开源溯源 : 无（clean-room 自研，未借鉴任何开源实现）
   输入契约 : adwData 待哈希数据 [1..32]；iLen 有效字数（自动钳位 0..32）
   输出契约 : 返回值 = 32 位哈希值；dwBytes 参与哈希的字节数；xValid 输入有效
   算法说明 : 逐字节 h += b；h += h<<10；h ^= h>>6。终混 h += h<<3；h ^= h>>11；h += h<<15
              全部移位量固定且小于 32 位宽
   修改记录 : v1.0.0 2026-11-24 初版
   =========================================================================== *)

FUNCTION FC_DL_HashJenkinsOneAtATime : DWORD
VAR_INPUT
    adwData : ARRAY[1..32] OF DWORD;   // 待哈希数据字 | data words to hash
    iLen : INT := 0;                   // 有效字数 0..32 | valid word count 0..32
END_VAR
VAR_OUTPUT
    dwBytes : DWORD;                   // 参与哈希的字节数 | hashed byte count
    xValid : BOOL;                     // 输入有效标志 | inputs valid flag
END_VAR
VAR
    dwHash : DWORD := 0;               // 哈希累加值 | hash accumulator
    dwByte : DWORD;                    // 当前字节 | current byte
    iN : INT;                          // 钳位后字数 | clamped word count
    i : INT;                           // 字下标 | word index
    b : INT;                           // 字节下标 0..3 | byte index 0..3
END_VAR

// ---- 输出预置 ----
dwBytes := 0;
xValid := FALSE;
FC_DL_HashJenkinsOneAtATime := 0;

// ---- 长度钳位 ----
iN := iLen;
IF iN < 0 THEN
    iN := 0;
ELSIF iN > 32 THEN
    iN := 32;
END_IF

// ---- 正文混合 ----
FOR i := 1 TO iN DO
    FOR b := 0 TO 3 DO
        dwByte := SHR(adwData[i], b * 8) AND 16#000000FF;
        dwHash := dwHash + dwByte;
        dwHash := dwHash + SHL(dwHash, 10);        // 左移 10 位，小于位宽
        dwHash := dwHash XOR SHR(dwHash, 6);       // 右移 6 位，小于位宽
    END_FOR
END_FOR

// ---- 终混：用于把末字节的影响扩散到全字 ----
dwHash := dwHash + SHL(dwHash, 3);
dwHash := dwHash XOR SHR(dwHash, 11);
dwHash := dwHash + SHL(dwHash, 15);

dwBytes := INT_TO_DWORD(iN) * INT_TO_DWORD(4);
xValid := TRUE;
FC_DL_HashJenkinsOneAtATime := dwHash;
END_FUNCTION

(* ---- FC_DL_HashMurmurLite.st ---- *)
(* ===========================================================================
   组件名   : FC_DL_HashMurmurLite
   分类     : DL_Algo / 哈希与完整性摘要
   一句话   : Murmur 简化版（不含尾部字节处理），含 32 位循环移位与终混雪崩
   复杂度   : 2        版本 : v1.0.0        日期 : 2026-11-24
   开源溯源 : 无（clean-room 自研，未借鉴任何开源实现）
   输入契约 : adwData 待哈希数据 [1..32]；iLen 有效字数（自动钳位 0..32）
              dwSeed 种子值
   输出契约 : 返回值 = 32 位哈希值；dwBytes 参与哈希的字节数；xValid 输入有效
   算法说明 : 循环左移用 SHL(x,n) OR SHR(x,32−n) 拼合实现，n 与 32−n 均小于 32；
              c1=16#CC9E2D51、c2=16#1B873593，终混取 16#85EBCA6B 与 16#C2B2AE35
              简化点：不处理非 4 字节整数倍的尾部，调用方须补齐零字节
   修改记录 : v1.0.0 2026-11-24 初版
   =========================================================================== *)

FUNCTION FC_DL_HashMurmurLite : DWORD
VAR_INPUT
    adwData : ARRAY[1..32] OF DWORD;   // 待哈希数据字 | data words to hash
    iLen : INT := 0;                   // 有效字数 0..32 | valid word count 0..32
    dwSeed : DWORD := 0;               // 哈希种子 | hash seed
END_VAR
VAR_OUTPUT
    dwBytes : DWORD;                   // 参与哈希的字节数 | hashed byte count
    xValid : BOOL;                     // 输入有效标志 | inputs valid flag
END_VAR
VAR
    dwH : DWORD;                       // 哈希累加值 | hash accumulator
    dwK : DWORD;                       // 单字混合值 | per word mix value
    iN : INT;                          // 钳位后字数 | clamped word count
    i : INT;                           // 字下标 | word index
END_VAR

// ---- 输出预置 ----
dwBytes := 0;
xValid := FALSE;
FC_DL_HashMurmurLite := 0;

// ---- 长度钳位 ----
iN := iLen;
IF iN < 0 THEN
    iN := 0;
ELSIF iN > 32 THEN
    iN := 32;
END_IF

dwH := dwSeed;

// ---- 正文：逐字混合 ----
FOR i := 1 TO iN DO
    dwK := adwData[i];
    dwK := dwK * 16#CC9E2D51;                      // 乘 c1
    dwK := SHL(dwK, 15) OR SHR(dwK, 17);           // 循环左移 15 位
    dwK := dwK * 16#1B873593;                      // 乘 c2

    dwH := dwH XOR dwK;
    dwH := SHL(dwH, 13) OR SHR(dwH, 19);           // 循环左移 13 位
    dwH := dwH * 5 + 16#E6546B64;
END_FOR

// ---- 长度混合：把字数折算成字节数并入哈希 ----
dwH := dwH XOR (INT_TO_DWORD(iN) * INT_TO_DWORD(4));

// ---- 终混：保证末位变化可扩散到全字 ----
dwH := dwH XOR SHR(dwH, 16);
dwH := dwH * 16#85EBCA6B;
dwH := dwH XOR SHR(dwH, 13);
dwH := dwH * 16#C2B2AE35;
dwH := dwH XOR SHR(dwH, 16);

dwBytes := INT_TO_DWORD(iN) * INT_TO_DWORD(4);
xValid := TRUE;
FC_DL_HashMurmurLite := dwH;
END_FUNCTION

(* ---- FC_DL_HashSdbmArray.st ---- *)
(* ===========================================================================
   组件名   : FC_DL_HashSdbmArray
   分类     : DL_Algo / 哈希与完整性摘要
   一句话   : sdbm 哈希，逐字节执行 h = b + (h<<6) + (h<<16) − h
   复杂度   : 1        版本 : v1.0.0        日期 : 2026-11-24
   开源溯源 : 无（clean-room 自研，未借鉴任何开源实现）
   输入契约 : adwData 待哈希数据 [1..32]；iLen 有效字数（自动钳位 0..32）
   输出契约 : 返回值 = 32 位哈希值；dwBytes 参与哈希的字节数；xValid 输入有效
   算法说明 : 移位量固定为 6 与 16，均小于 32 位宽，不触发未定义移位
   修改记录 : v1.0.0 2026-11-24 初版
   =========================================================================== *)

FUNCTION FC_DL_HashSdbmArray : DWORD
VAR_INPUT
    adwData : ARRAY[1..32] OF DWORD;   // 待哈希数据字 | data words to hash
    iLen : INT := 0;                   // 有效字数 0..32 | valid word count 0..32
END_VAR
VAR_OUTPUT
    dwBytes : DWORD;                   // 参与哈希的字节数 | hashed byte count
    xValid : BOOL;                     // 输入有效标志 | inputs valid flag
END_VAR
VAR
    dwHash : DWORD := 0;               // sdbm 累加值 | sdbm accumulator
    dwByte : DWORD;                    // 当前字节 | current byte
    iN : INT;                          // 钳位后字数 | clamped word count
    i : INT;                           // 字下标 | word index
    b : INT;                           // 字节下标 0..3 | byte index 0..3
END_VAR

// ---- 输出预置 ----
dwBytes := 0;
xValid := FALSE;
FC_DL_HashSdbmArray := 0;

// ---- 长度钳位 ----
iN := iLen;
IF iN < 0 THEN
    iN := 0;
ELSIF iN > 32 THEN
    iN := 32;
END_IF

// ---- 逐字逐字节处理 ----
FOR i := 1 TO iN DO
    FOR b := 0 TO 3 DO
        dwByte := SHR(adwData[i], b * 8) AND 16#000000FF;
        dwHash := dwByte + SHL(dwHash, 6) + SHL(dwHash, 16) - dwHash;
    END_FOR
END_FOR

dwBytes := INT_TO_DWORD(iN) * INT_TO_DWORD(4);
xValid := TRUE;
FC_DL_HashSdbmArray := dwHash;
END_FUNCTION

(* ---- FC_DL_HashXorFold.st ---- *)
(* ===========================================================================
   组件名   : FC_DL_HashXorFold
   分类     : DL_Algo / 哈希与完整性摘要
   一句话   : 异或折叠哈希：先把每个 DWORD 的四字节折叠成单字节，再与累加值混合
   复杂度   : 1        版本 : v1.0.0        日期 : 2026-11-24
   开源溯源 : 无（clean-room 自研，未借鉴任何开源实现）
   输入契约 : adwData 待哈希数据 [1..32]；iLen 有效字数（自动钳位 0..32）
   输出契约 : 返回值 = 32 位哈希值；dwBytes 参与哈希的字节数；xValid 输入有效
   算法说明 : fold = b0^b1^b2^b3；h = (h ^ fold) * 16#01000193；h = h ^ (h>>13)
              折叠保留了各字节奇偶信息，混合步保证低位扩散
   修改记录 : v1.0.0 2026-11-24 初版
   =========================================================================== *)

FUNCTION FC_DL_HashXorFold : DWORD
VAR_INPUT
    adwData : ARRAY[1..32] OF DWORD;   // 待哈希数据字 | data words to hash
    iLen : INT := 0;                   // 有效字数 0..32 | valid word count 0..32
END_VAR
VAR_OUTPUT
    dwBytes : DWORD;                   // 参与哈希的字节数 | hashed byte count
    xValid : BOOL;                     // 输入有效标志 | inputs valid flag
END_VAR
VAR
    dwHash : DWORD := 16#811C9DC5;     // 哈希累加值 | hash accumulator
    dwFold : DWORD;                    // 单字折叠值 | folded byte of one word
    dwByte : DWORD;                    // 当前字节 | current byte
    iN : INT;                          // 钳位后字数 | clamped word count
    i : INT;                           // 字下标 | word index
    b : INT;                           // 字节下标 0..3 | byte index 0..3
END_VAR

// ---- 输出预置 ----
dwBytes := 0;
xValid := FALSE;
FC_DL_HashXorFold := 16#811C9DC5;

// ---- 长度钳位 ----
iN := iLen;
IF iN < 0 THEN
    iN := 0;
ELSIF iN > 32 THEN
    iN := 32;
END_IF

// ---- 折叠 + 混合 ----
FOR i := 1 TO iN DO
    dwFold := 0;
    FOR b := 0 TO 3 DO
        dwByte := SHR(adwData[i], b * 8) AND 16#000000FF;
        dwFold := dwFold XOR dwByte;               // 四字节异或折叠
    END_FOR
    dwHash := (dwHash XOR dwFold) * 16#01000193;   // 与折叠值混合
    dwHash := dwHash XOR SHR(dwHash, 13);          // 高位回灌低位
END_FOR

dwBytes := INT_TO_DWORD(iN) * INT_TO_DWORD(4);
xValid := TRUE;
FC_DL_HashXorFold := dwHash;
END_FUNCTION

(* ---- FC_DL_HoneStonePressureCalc.st ---- *)
(*
  DL Factory R88 | FC_DL_HoneStonePressureCalc
  功能：算珩磨油石比压 p=F/(n·L·W)，N/mm² 按 ×10 换算为 bar，并按工艺带宽判合格
  开源溯源：无（clean-room 自研，依据公开工艺公式 接触比压定义式 p=F/A，许可证=MIT，借鉴点=公式结构）
  规则：R1-R16 全遵守；R88 简单件标量形（纯标量入参出参，无循环体、无方法、无属性、无数组）
*)
FUNCTION FC_DL_HoneStonePressureCalc : REAL
VAR_INPUT
    fForceN : REAL := 1200.0; // 油石总法向压紧力 F [N] / total normal stone force [N]
    nStoneCount : DINT := 6; // 油石条数 n（整数入参，无 NaN 可能） [条] / number of stones [-]
    fStoneLengthMm : REAL := 100.0; // 单条油石接触长度 L [mm] / stone contact length [mm]
    fStoneWidthMm : REAL := 10.0; // 单条油石接触宽度 W [mm] / stone contact width [mm]
    fMinBar : REAL := 2.0; // 比压允许下限（工艺带宽） [bar] / lower pressure band [bar]
    fMaxBar : REAL := 8.0; // 比压允许上限（工艺带宽） [bar] / upper pressure band [bar]
END_VAR
VAR_OUTPUT
    fPressBar : REAL; // 油石比压 p（N/mm²×10） [bar] / stone specific pressure [bar]
    xInBand : BOOL; // TRUE=比压落在允许带宽内 [-] / TRUE when inside the band [-]
END_VAR
VAR
    fStones : REAL; // 油石条数实数化 [-] / stone count as real [-]
    fAreaTotalMm2 : REAL; // 总接触面积 n·L·W（除零判据） [mm²] / total contact area, the divisor [mm^2]
    fPressMpa : REAL; // 比压 N/mm²（数值等同 MPa） [N/mm²] / specific pressure [N/mm^2]
END_VAR

// 段 1｜出口预置
FC_DL_HoneStonePressureCalc := -1.0; // 哨兵返回 -1（无效） [-] / sentinel return -1, invalid [-]
fPressBar := 0.0; // 比压预置零 [bar] / pressure preset zero [bar]
xInBand := FALSE; // 带宽位预置 FALSE（未判定前不认合格） [-] / band flag preset false [-]

// 段 2｜非有限拦截 + 域闸
IF NOT (fForceN > -1.0E30 AND fForceN < 1.0E30) OR NOT (fStoneLengthMm > -1.0E30 AND fStoneLengthMm < 1.0E30) OR NOT (fStoneWidthMm > -1.0E30 AND fStoneWidthMm < 1.0E30) THEN
    RETURN; // 压紧力/油石长宽任一非有限即拒算 [-] / any non finite input rejected [-]
END_IF
IF NOT (fMinBar > -1.0E30 AND fMinBar < 1.0E30) OR NOT (fMaxBar > -1.0E30 AND fMaxBar < 1.0E30) THEN
    RETURN; // 带宽上下限任一非有限则判据静默失效，故先拦 [bar] / band limits must be finite [bar]
END_IF
IF fForceN < 0.0 OR fStoneLengthMm < 1.0E-9 OR fStoneWidthMm < 1.0E-9 THEN
    RETURN; // 力非负闸 + 长宽正域闸（分母不得为零） [N, mm] / non negative force and positive geometry [N, mm]
END_IF
IF nStoneCount < 1 OR fMinBar <= 0.0 OR fMaxBar <= fMinBar THEN
    RETURN; // 条数下限闸 + 带宽自洽闸（整数域无 NaN 可能） [条, bar] / count and band gates
END_IF

// 段 3｜计算
fStones := DINT_TO_REAL(nStoneCount); // DINT→REAL 标准转换函数（R10） [-] / standard conversion (R10) [-]
fAreaTotalMm2 := fStones * fStoneLengthMm * fStoneWidthMm; // 无量纲 × mm × mm = mm²，A=n·L·W [mm²] / [mm^2]
IF fAreaTotalMm2 < 1.0E-9 THEN
    RETURN; // 除法前分母闸：总面积必须大于 1E-9 才可作除数 [mm²] / denominator gate [mm^2]
END_IF
fPressMpa := fForceN / fAreaTotalMm2; // N ÷ mm² = N/mm²（数值等同 MPa） [N/mm²] / [N] / [mm^2] = [N/mm^2]
fPressBar := fPressMpa * 10.0; // 1 N/mm² = 1 MPa = 10 bar，故 ×10 换算 [bar] / 1 MPa equals 10 bar [bar]

// 段 4｜判定与饱和
IF NOT (fPressBar > -1.0E30 AND fPressBar < 1.0E30) THEN
    RETURN; // 结果非有限再拦一次 [-] / re-check the result for finiteness [-]
END_IF
xInBand := (fPressBar >= fMinBar) AND (fPressBar <= fMaxBar); // 双侧闭区间直比 [bar] / closed two sided band compare [bar]

// 段 5｜出口自检
IF fPressBar < 0.0 THEN
    RETURN; // 出口自检：比压不得为负（负值说明力符号错） [bar] / pressure must not be negative [bar]
END_IF
FC_DL_HoneStonePressureCalc := fPressBar; // 返回油石比压 [bar] / return the stone specific pressure [bar]
END_FUNCTION
